REGION Network 25: Level Conveyors Tower 1 - SYSTEM 2
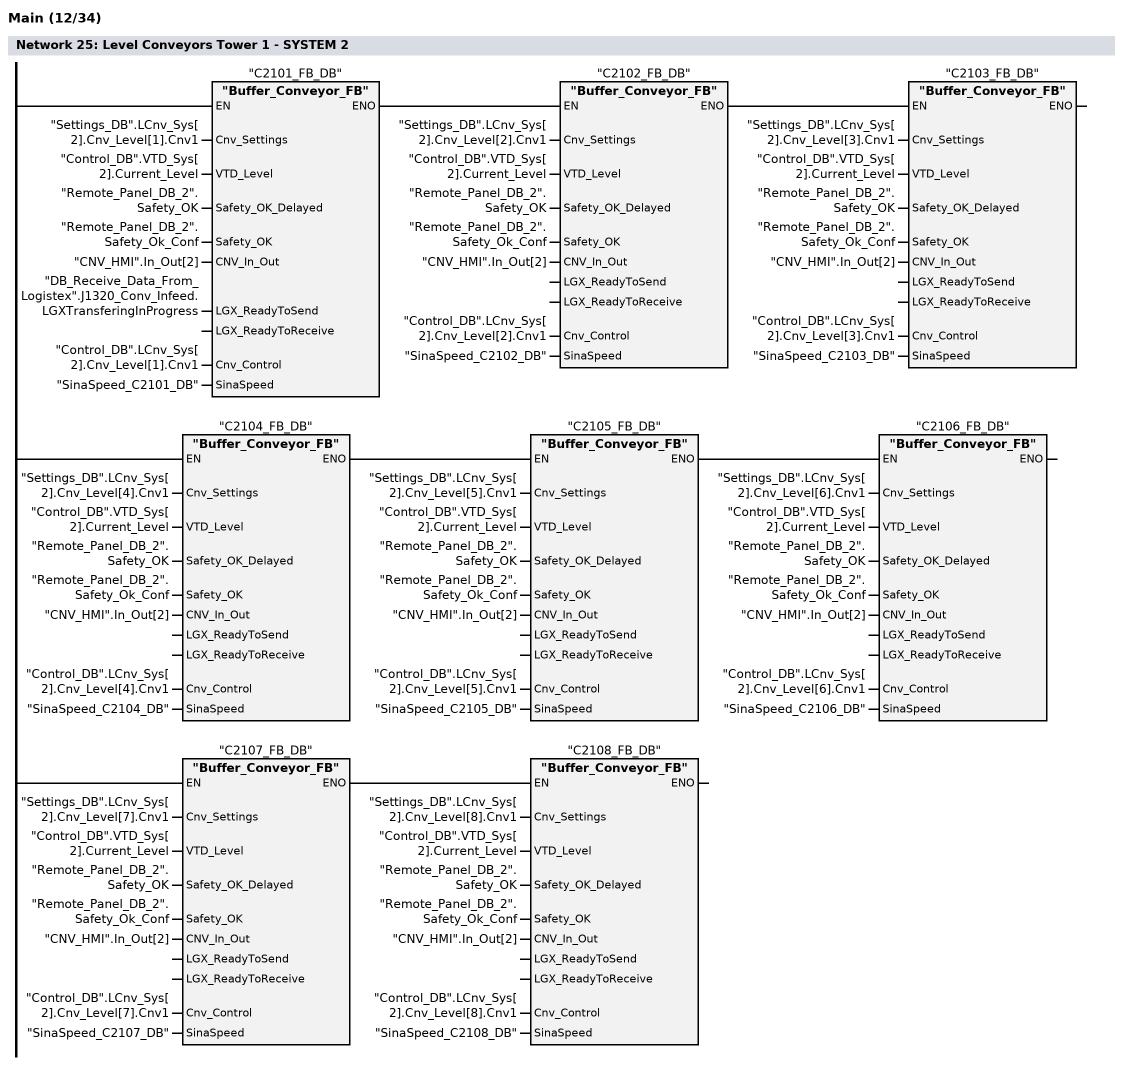
   RUNG wire#powerrail
      "C2101_FB_DB"(Cnv_Settings := "Settings_DB".LCnv_Sys[2].Cnv_Level[1].Cnv1, VTD_Level := "Control_DB".VTD_Sys[2].Current_Level, Safety_OK_Delayed := "Remote_Panel_DB_2".Safety_OK, Safety_OK := "Remote_Panel_DB_2".Safety_Ok_Conf, CNV_In_Out := "CNV_HMI".In_Out[2], LGX_ReadyToSend := "DB_Receive_Data_From_Logistex".J1320_Conv_Infeed.LGXTransferingInProgress, LGX_ReadyToReceive :=, Cnv_Control := "Control_DB".LCnv_Sys[2].Cnv_Level[1].Cnv1, SinaSpeed := "SinaSpeed_C2101_DB")
      "C2102_FB_DB"(Cnv_Settings := "Settings_DB".LCnv_Sys[2].Cnv_Level[2].Cnv1, VTD_Level := "Control_DB".VTD_Sys[2].Current_Level, Safety_OK_Delayed := "Remote_Panel_DB_2".Safety_OK, Safety_OK := "Remote_Panel_DB_2".Safety_Ok_Conf, CNV_In_Out := "CNV_HMI".In_Out[2], LGX_ReadyToSend :=, LGX_ReadyToReceive :=, Cnv_Control := "Control_DB".LCnv_Sys[2].Cnv_Level[2].Cnv1, SinaSpeed := "SinaSpeed_C2102_DB")
      "C2103_FB_DB"(Cnv_Settings := "Settings_DB".LCnv_Sys[2].Cnv_Level[3].Cnv1, VTD_Level := "Control_DB".VTD_Sys[2].Current_Level, Safety_OK_Delayed := "Remote_Panel_DB_2".Safety_OK, Safety_OK := "Remote_Panel_DB_2".Safety_Ok_Conf, CNV_In_Out := "CNV_HMI".In_Out[2], LGX_ReadyToSend :=, LGX_ReadyToReceive :=, Cnv_Control := "Control_DB".LCnv_Sys[2].Cnv_Level[3].Cnv1, SinaSpeed := "SinaSpeed_C2103_DB")
   END_RUNG
   RUNG wire#powerrail
      "C2104_FB_DB"(Cnv_Settings := "Settings_DB".LCnv_Sys[2].Cnv_Level[4].Cnv1, VTD_Level := "Control_DB".VTD_Sys[2].Current_Level, Safety_OK_Delayed := "Remote_Panel_DB_2".Safety_OK, Safety_OK := "Remote_Panel_DB_2".Safety_Ok_Conf, CNV_In_Out := "CNV_HMI".In_Out[2], LGX_ReadyToSend :=, LGX_ReadyToReceive :=, Cnv_Control := "Control_DB".LCnv_Sys[2].Cnv_Level[4].Cnv1, SinaSpeed := "SinaSpeed_C2104_DB")
      "C2105_FB_DB"(Cnv_Settings := "Settings_DB".LCnv_Sys[2].Cnv_Level[5].Cnv1, VTD_Level := "Control_DB".VTD_Sys[2].Current_Level, Safety_OK_Delayed := "Remote_Panel_DB_2".Safety_OK, Safety_OK := "Remote_Panel_DB_2".Safety_Ok_Conf, CNV_In_Out := "CNV_HMI".In_Out[2], LGX_ReadyToSend :=, LGX_ReadyToReceive :=, Cnv_Control := "Control_DB".LCnv_Sys[2].Cnv_Level[5].Cnv1, SinaSpeed := "SinaSpeed_C2105_DB")
      "C2106_FB_DB"(Cnv_Settings := "Settings_DB".LCnv_Sys[2].Cnv_Level[6].Cnv1, VTD_Level := "Control_DB".VTD_Sys[2].Current_Level, Safety_OK_Delayed := "Remote_Panel_DB_2".Safety_OK, Safety_OK := "Remote_Panel_DB_2".Safety_Ok_Conf, CNV_In_Out := "CNV_HMI".In_Out[2], LGX_ReadyToSend :=, LGX_ReadyToReceive :=, Cnv_Control := "Control_DB".LCnv_Sys[2].Cnv_Level[6].Cnv1, SinaSpeed := "SinaSpeed_C2106_DB")
   END_RUNG
   RUNG wire#powerrail
      "C2107_FB_DB"(Cnv_Settings := "Settings_DB".LCnv_Sys[2].Cnv_Level[7].Cnv1, VTD_Level := "Control_DB".VTD_Sys[2].Current_Level, Safety_OK_Delayed := "Remote_Panel_DB_2".Safety_OK, Safety_OK := "Remote_Panel_DB_2".Safety_Ok_Conf, CNV_In_Out := "CNV_HMI".In_Out[2], LGX_ReadyToSend :=, LGX_ReadyToReceive :=, Cnv_Control := "Control_DB".LCnv_Sys[2].Cnv_Level[7].Cnv1, SinaSpeed := "SinaSpeed_C2107_DB")
      "C2108_FB_DB"(Cnv_Settings := "Settings_DB".LCnv_Sys[2].Cnv_Level[8].Cnv1, VTD_Level := "Control_DB".VTD_Sys[2].Current_Level, Safety_OK_Delayed := "Remote_Panel_DB_2".Safety_OK, Safety_OK := "Remote_Panel_DB_2".Safety_Ok_Conf, CNV_In_Out := "CNV_HMI".In_Out[2], LGX_ReadyToSend :=, LGX_ReadyToReceive :=, Cnv_Control := "Control_DB".LCnv_Sys[2].Cnv_Level[8].Cnv1, SinaSpeed := "SinaSpeed_C2108_DB")
   END_RUNG
   // the same network as SCL:
   "C2101_FB_DB"(Cnv_Settings := "Settings_DB".LCnv_Sys[2].Cnv_Level[1].Cnv1,   // "Buffer_Conveyor_FB"
                 VTD_Level := "Control_DB".VTD_Sys[2].Current_Level,
                 Safety_OK_Delayed := "Remote_Panel_DB_2".Safety_OK,
                 Safety_OK := "Remote_Panel_DB_2".Safety_Ok_Conf,
                 CNV_In_Out := "CNV_HMI".In_Out[2],
                 LGX_ReadyToSend := "DB_Receive_Data_From_Logistex".J1320_Conv_Infeed.LGXTransferingInProgress,
                 Cnv_Control := "Control_DB".LCnv_Sys[2].Cnv_Level[1].Cnv1,
                 SinaSpeed := "SinaSpeed_C2101_DB",
                 ENO => #_w1);
   "C2102_FB_DB"(EN := #_w1,   // "Buffer_Conveyor_FB"
                 Cnv_Settings := "Settings_DB".LCnv_Sys[2].Cnv_Level[2].Cnv1,
                 VTD_Level := "Control_DB".VTD_Sys[2].Current_Level,
                 Safety_OK_Delayed := "Remote_Panel_DB_2".Safety_OK,
                 Safety_OK := "Remote_Panel_DB_2".Safety_Ok_Conf,
                 CNV_In_Out := "CNV_HMI".In_Out[2],
                 Cnv_Control := "Control_DB".LCnv_Sys[2].Cnv_Level[2].Cnv1,
                 SinaSpeed := "SinaSpeed_C2102_DB",
                 ENO => #_w2);
   IF #_w2 THEN
       "C2103_FB_DB"(Cnv_Settings := "Settings_DB".LCnv_Sys[2].Cnv_Level[3].Cnv1,   // "Buffer_Conveyor_FB"
                     VTD_Level := "Control_DB".VTD_Sys[2].Current_Level,
                     Safety_OK_Delayed := "Remote_Panel_DB_2".Safety_OK,
                     Safety_OK := "Remote_Panel_DB_2".Safety_Ok_Conf,
                     CNV_In_Out := "CNV_HMI".In_Out[2],
                     Cnv_Control := "Control_DB".LCnv_Sys[2].Cnv_Level[3].Cnv1,
                     SinaSpeed := "SinaSpeed_C2103_DB");
   END_IF;
   "C2104_FB_DB"(Cnv_Settings := "Settings_DB".LCnv_Sys[2].Cnv_Level[4].Cnv1,   // "Buffer_Conveyor_FB"
                 VTD_Level := "Control_DB".VTD_Sys[2].Current_Level,
                 Safety_OK_Delayed := "Remote_Panel_DB_2".Safety_OK,
                 Safety_OK := "Remote_Panel_DB_2".Safety_Ok_Conf,
                 CNV_In_Out := "CNV_HMI".In_Out[2],
                 Cnv_Control := "Control_DB".LCnv_Sys[2].Cnv_Level[4].Cnv1,
                 SinaSpeed := "SinaSpeed_C2104_DB",
                 ENO => #_w3);
   "C2105_FB_DB"(EN := #_w3,   // "Buffer_Conveyor_FB"
                 Cnv_Settings := "Settings_DB".LCnv_Sys[2].Cnv_Level[5].Cnv1,
                 VTD_Level := "Control_DB".VTD_Sys[2].Current_Level,
                 Safety_OK_Delayed := "Remote_Panel_DB_2".Safety_OK,
                 Safety_OK := "Remote_Panel_DB_2".Safety_Ok_Conf,
                 CNV_In_Out := "CNV_HMI".In_Out[2],
                 Cnv_Control := "Control_DB".LCnv_Sys[2].Cnv_Level[5].Cnv1,
                 SinaSpeed := "SinaSpeed_C2105_DB",
                 ENO => #_w4);
   IF #_w4 THEN
       "C2106_FB_DB"(Cnv_Settings := "Settings_DB".LCnv_Sys[2].Cnv_Level[6].Cnv1,   // "Buffer_Conveyor_FB"
                     VTD_Level := "Control_DB".VTD_Sys[2].Current_Level,
                     Safety_OK_Delayed := "Remote_Panel_DB_2".Safety_OK,
                     Safety_OK := "Remote_Panel_DB_2".Safety_Ok_Conf,
                     CNV_In_Out := "CNV_HMI".In_Out[2],
                     Cnv_Control := "Control_DB".LCnv_Sys[2].Cnv_Level[6].Cnv1,
                     SinaSpeed := "SinaSpeed_C2106_DB");
   END_IF;
   "C2107_FB_DB"(Cnv_Settings := "Settings_DB".LCnv_Sys[2].Cnv_Level[7].Cnv1,   // "Buffer_Conveyor_FB"
                 VTD_Level := "Control_DB".VTD_Sys[2].Current_Level,
                 Safety_OK_Delayed := "Remote_Panel_DB_2".Safety_OK,
                 Safety_OK := "Remote_Panel_DB_2".Safety_Ok_Conf,
                 CNV_In_Out := "CNV_HMI".In_Out[2],
                 Cnv_Control := "Control_DB".LCnv_Sys[2].Cnv_Level[7].Cnv1,
                 SinaSpeed := "SinaSpeed_C2107_DB",
                 ENO => #_w5);
   IF #_w5 THEN
       "C2108_FB_DB"(Cnv_Settings := "Settings_DB".LCnv_Sys[2].Cnv_Level[8].Cnv1,   // "Buffer_Conveyor_FB"
                     VTD_Level := "Control_DB".VTD_Sys[2].Current_Level,
                     Safety_OK_Delayed := "Remote_Panel_DB_2".Safety_OK,
                     Safety_OK := "Remote_Panel_DB_2".Safety_Ok_Conf,
                     CNV_In_Out := "CNV_HMI".In_Out[2],
                     Cnv_Control := "Control_DB".LCnv_Sys[2].Cnv_Level[8].Cnv1,
                     SinaSpeed := "SinaSpeed_C2108_DB");
   END_IF;
END_REGION

REGION Network 26: Level Conveyors Tower 2 - SYSTEM 2
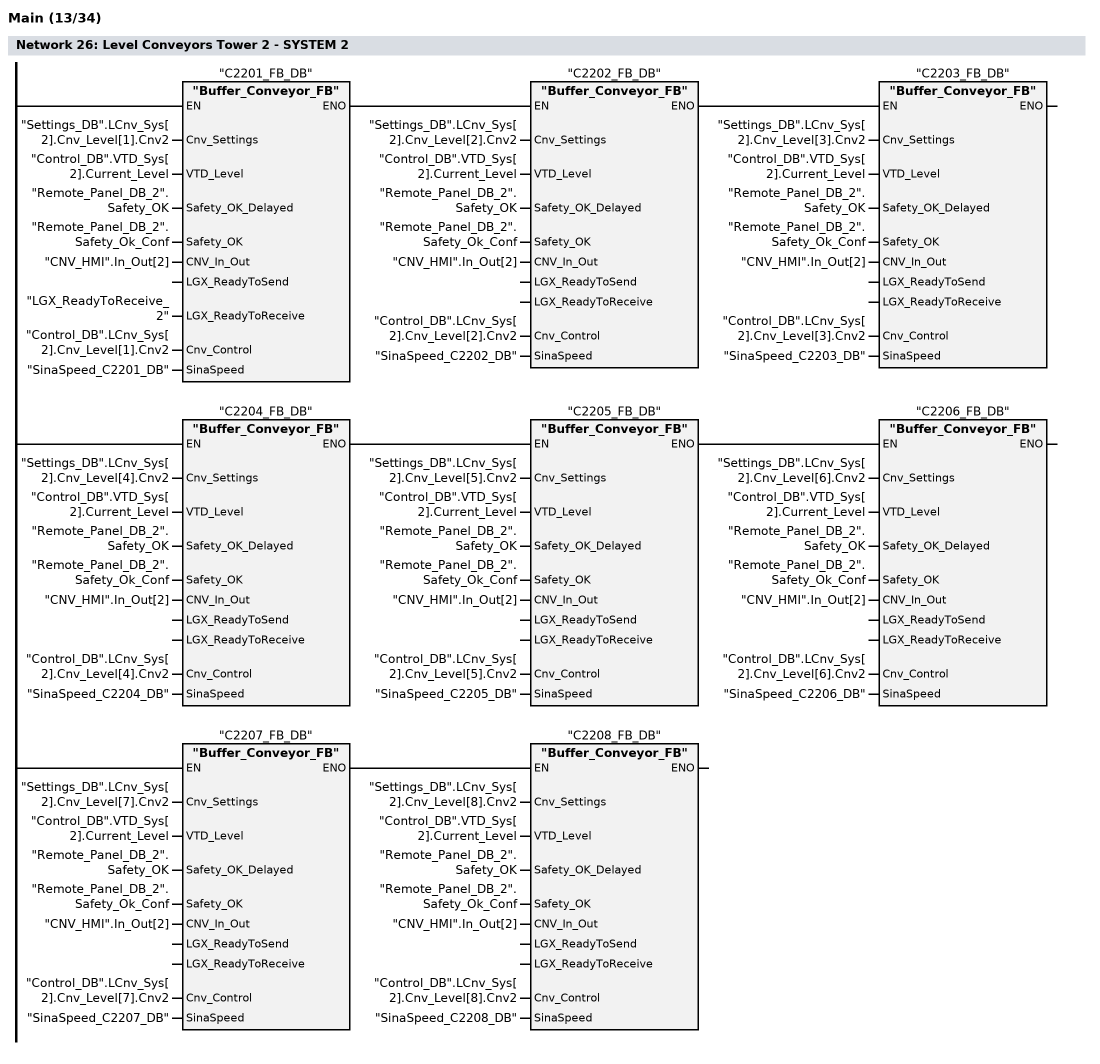
   RUNG wire#powerrail
      "C2201_FB_DB"(Cnv_Settings := "Settings_DB".LCnv_Sys[2].Cnv_Level[1].Cnv2, VTD_Level := "Control_DB".VTD_Sys[2].Current_Level, Safety_OK_Delayed := "Remote_Panel_DB_2".Safety_OK, Safety_OK := "Remote_Panel_DB_2".Safety_Ok_Conf, CNV_In_Out := "CNV_HMI".In_Out[2], LGX_ReadyToSend :=, LGX_ReadyToReceive := "LGX_ReadyToReceive_2", Cnv_Control := "Control_DB".LCnv_Sys[2].Cnv_Level[1].Cnv2, SinaSpeed := "SinaSpeed_C2201_DB")
      "C2202_FB_DB"(Cnv_Settings := "Settings_DB".LCnv_Sys[2].Cnv_Level[2].Cnv2, VTD_Level := "Control_DB".VTD_Sys[2].Current_Level, Safety_OK_Delayed := "Remote_Panel_DB_2".Safety_OK, Safety_OK := "Remote_Panel_DB_2".Safety_Ok_Conf, CNV_In_Out := "CNV_HMI".In_Out[2], LGX_ReadyToSend :=, LGX_ReadyToReceive :=, Cnv_Control := "Control_DB".LCnv_Sys[2].Cnv_Level[2].Cnv2, SinaSpeed := "SinaSpeed_C2202_DB")
      "C2203_FB_DB"(Cnv_Settings := "Settings_DB".LCnv_Sys[2].Cnv_Level[3].Cnv2, VTD_Level := "Control_DB".VTD_Sys[2].Current_Level, Safety_OK_Delayed := "Remote_Panel_DB_2".Safety_OK, Safety_OK := "Remote_Panel_DB_2".Safety_Ok_Conf, CNV_In_Out := "CNV_HMI".In_Out[2], LGX_ReadyToSend :=, LGX_ReadyToReceive :=, Cnv_Control := "Control_DB".LCnv_Sys[2].Cnv_Level[3].Cnv2, SinaSpeed := "SinaSpeed_C2203_DB")
   END_RUNG
   RUNG wire#powerrail
      "C2204_FB_DB"(Cnv_Settings := "Settings_DB".LCnv_Sys[2].Cnv_Level[4].Cnv2, VTD_Level := "Control_DB".VTD_Sys[2].Current_Level, Safety_OK_Delayed := "Remote_Panel_DB_2".Safety_OK, Safety_OK := "Remote_Panel_DB_2".Safety_Ok_Conf, CNV_In_Out := "CNV_HMI".In_Out[2], LGX_ReadyToSend :=, LGX_ReadyToReceive :=, Cnv_Control := "Control_DB".LCnv_Sys[2].Cnv_Level[4].Cnv2, SinaSpeed := "SinaSpeed_C2204_DB")
      "C2205_FB_DB"(Cnv_Settings := "Settings_DB".LCnv_Sys[2].Cnv_Level[5].Cnv2, VTD_Level := "Control_DB".VTD_Sys[2].Current_Level, Safety_OK_Delayed := "Remote_Panel_DB_2".Safety_OK, Safety_OK := "Remote_Panel_DB_2".Safety_Ok_Conf, CNV_In_Out := "CNV_HMI".In_Out[2], LGX_ReadyToSend :=, LGX_ReadyToReceive :=, Cnv_Control := "Control_DB".LCnv_Sys[2].Cnv_Level[5].Cnv2, SinaSpeed := "SinaSpeed_C2205_DB")
      "C2206_FB_DB"(Cnv_Settings := "Settings_DB".LCnv_Sys[2].Cnv_Level[6].Cnv2, VTD_Level := "Control_DB".VTD_Sys[2].Current_Level, Safety_OK_Delayed := "Remote_Panel_DB_2".Safety_OK, Safety_OK := "Remote_Panel_DB_2".Safety_Ok_Conf, CNV_In_Out := "CNV_HMI".In_Out[2], LGX_ReadyToSend :=, LGX_ReadyToReceive :=, Cnv_Control := "Control_DB".LCnv_Sys[2].Cnv_Level[6].Cnv2, SinaSpeed := "SinaSpeed_C2206_DB")
   END_RUNG
   RUNG wire#powerrail
      "C2207_FB_DB"(Cnv_Settings := "Settings_DB".LCnv_Sys[2].Cnv_Level[7].Cnv2, VTD_Level := "Control_DB".VTD_Sys[2].Current_Level, Safety_OK_Delayed := "Remote_Panel_DB_2".Safety_OK, Safety_OK := "Remote_Panel_DB_2".Safety_Ok_Conf, CNV_In_Out := "CNV_HMI".In_Out[2], LGX_ReadyToSend :=, LGX_ReadyToReceive :=, Cnv_Control := "Control_DB".LCnv_Sys[2].Cnv_Level[7].Cnv2, SinaSpeed := "SinaSpeed_C2207_DB")
      "C2208_FB_DB"(Cnv_Settings := "Settings_DB".LCnv_Sys[2].Cnv_Level[8].Cnv2, VTD_Level := "Control_DB".VTD_Sys[2].Current_Level, Safety_OK_Delayed := "Remote_Panel_DB_2".Safety_OK, Safety_OK := "Remote_Panel_DB_2".Safety_Ok_Conf, CNV_In_Out := "CNV_HMI".In_Out[2], LGX_ReadyToSend :=, LGX_ReadyToReceive :=, Cnv_Control := "Control_DB".LCnv_Sys[2].Cnv_Level[8].Cnv2, SinaSpeed := "SinaSpeed_C2208_DB")
   END_RUNG
   // the same network as SCL:
   "C2201_FB_DB"(Cnv_Settings := "Settings_DB".LCnv_Sys[2].Cnv_Level[1].Cnv2,   // "Buffer_Conveyor_FB"
                 VTD_Level := "Control_DB".VTD_Sys[2].Current_Level,
                 Safety_OK_Delayed := "Remote_Panel_DB_2".Safety_OK,
                 Safety_OK := "Remote_Panel_DB_2".Safety_Ok_Conf,
                 CNV_In_Out := "CNV_HMI".In_Out[2],
                 LGX_ReadyToReceive := "LGX_ReadyToReceive_2",
                 Cnv_Control := "Control_DB".LCnv_Sys[2].Cnv_Level[1].Cnv2,
                 SinaSpeed := "SinaSpeed_C2201_DB",
                 ENO => #_w1);
   "C2202_FB_DB"(EN := #_w1,   // "Buffer_Conveyor_FB"
                 Cnv_Settings := "Settings_DB".LCnv_Sys[2].Cnv_Level[2].Cnv2,
                 VTD_Level := "Control_DB".VTD_Sys[2].Current_Level,
                 Safety_OK_Delayed := "Remote_Panel_DB_2".Safety_OK,
                 Safety_OK := "Remote_Panel_DB_2".Safety_Ok_Conf,
                 CNV_In_Out := "CNV_HMI".In_Out[2],
                 Cnv_Control := "Control_DB".LCnv_Sys[2].Cnv_Level[2].Cnv2,
                 SinaSpeed := "SinaSpeed_C2202_DB",
                 ENO => #_w2);
   IF #_w2 THEN
       "C2203_FB_DB"(Cnv_Settings := "Settings_DB".LCnv_Sys[2].Cnv_Level[3].Cnv2,   // "Buffer_Conveyor_FB"
                     VTD_Level := "Control_DB".VTD_Sys[2].Current_Level,
                     Safety_OK_Delayed := "Remote_Panel_DB_2".Safety_OK,
                     Safety_OK := "Remote_Panel_DB_2".Safety_Ok_Conf,
                     CNV_In_Out := "CNV_HMI".In_Out[2],
                     Cnv_Control := "Control_DB".LCnv_Sys[2].Cnv_Level[3].Cnv2,
                     SinaSpeed := "SinaSpeed_C2203_DB");
   END_IF;
   "C2204_FB_DB"(Cnv_Settings := "Settings_DB".LCnv_Sys[2].Cnv_Level[4].Cnv2,   // "Buffer_Conveyor_FB"
                 VTD_Level := "Control_DB".VTD_Sys[2].Current_Level,
                 Safety_OK_Delayed := "Remote_Panel_DB_2".Safety_OK,
                 Safety_OK := "Remote_Panel_DB_2".Safety_Ok_Conf,
                 CNV_In_Out := "CNV_HMI".In_Out[2],
                 Cnv_Control := "Control_DB".LCnv_Sys[2].Cnv_Level[4].Cnv2,
                 SinaSpeed := "SinaSpeed_C2204_DB",
                 ENO => #_w3);
   "C2205_FB_DB"(EN := #_w3,   // "Buffer_Conveyor_FB"
                 Cnv_Settings := "Settings_DB".LCnv_Sys[2].Cnv_Level[5].Cnv2,
                 VTD_Level := "Control_DB".VTD_Sys[2].Current_Level,
                 Safety_OK_Delayed := "Remote_Panel_DB_2".Safety_OK,
                 Safety_OK := "Remote_Panel_DB_2".Safety_Ok_Conf,
                 CNV_In_Out := "CNV_HMI".In_Out[2],
                 Cnv_Control := "Control_DB".LCnv_Sys[2].Cnv_Level[5].Cnv2,
                 SinaSpeed := "SinaSpeed_C2205_DB",
                 ENO => #_w4);
   IF #_w4 THEN
       "C2206_FB_DB"(Cnv_Settings := "Settings_DB".LCnv_Sys[2].Cnv_Level[6].Cnv2,   // "Buffer_Conveyor_FB"
                     VTD_Level := "Control_DB".VTD_Sys[2].Current_Level,
                     Safety_OK_Delayed := "Remote_Panel_DB_2".Safety_OK,
                     Safety_OK := "Remote_Panel_DB_2".Safety_Ok_Conf,
                     CNV_In_Out := "CNV_HMI".In_Out[2],
                     Cnv_Control := "Control_DB".LCnv_Sys[2].Cnv_Level[6].Cnv2,
                     SinaSpeed := "SinaSpeed_C2206_DB");
   END_IF;
   "C2207_FB_DB"(Cnv_Settings := "Settings_DB".LCnv_Sys[2].Cnv_Level[7].Cnv2,   // "Buffer_Conveyor_FB"
                 VTD_Level := "Control_DB".VTD_Sys[2].Current_Level,
                 Safety_OK_Delayed := "Remote_Panel_DB_2".Safety_OK,
                 Safety_OK := "Remote_Panel_DB_2".Safety_Ok_Conf,
                 CNV_In_Out := "CNV_HMI".In_Out[2],
                 Cnv_Control := "Control_DB".LCnv_Sys[2].Cnv_Level[7].Cnv2,
                 SinaSpeed := "SinaSpeed_C2207_DB",
                 ENO => #_w5);
   IF #_w5 THEN
       "C2208_FB_DB"(Cnv_Settings := "Settings_DB".LCnv_Sys[2].Cnv_Level[8].Cnv2,   // "Buffer_Conveyor_FB"
                     VTD_Level := "Control_DB".VTD_Sys[2].Current_Level,
                     Safety_OK_Delayed := "Remote_Panel_DB_2".Safety_OK,
                     Safety_OK := "Remote_Panel_DB_2".Safety_Ok_Conf,
                     CNV_In_Out := "CNV_HMI".In_Out[2],
                     Cnv_Control := "Control_DB".LCnv_Sys[2].Cnv_Level[8].Cnv2,
                     SinaSpeed := "SinaSpeed_C2208_DB");
   END_IF;
END_REGION

REGION Network 27: SAFETY STOPPERS Tower 1 - SYSTEM 2
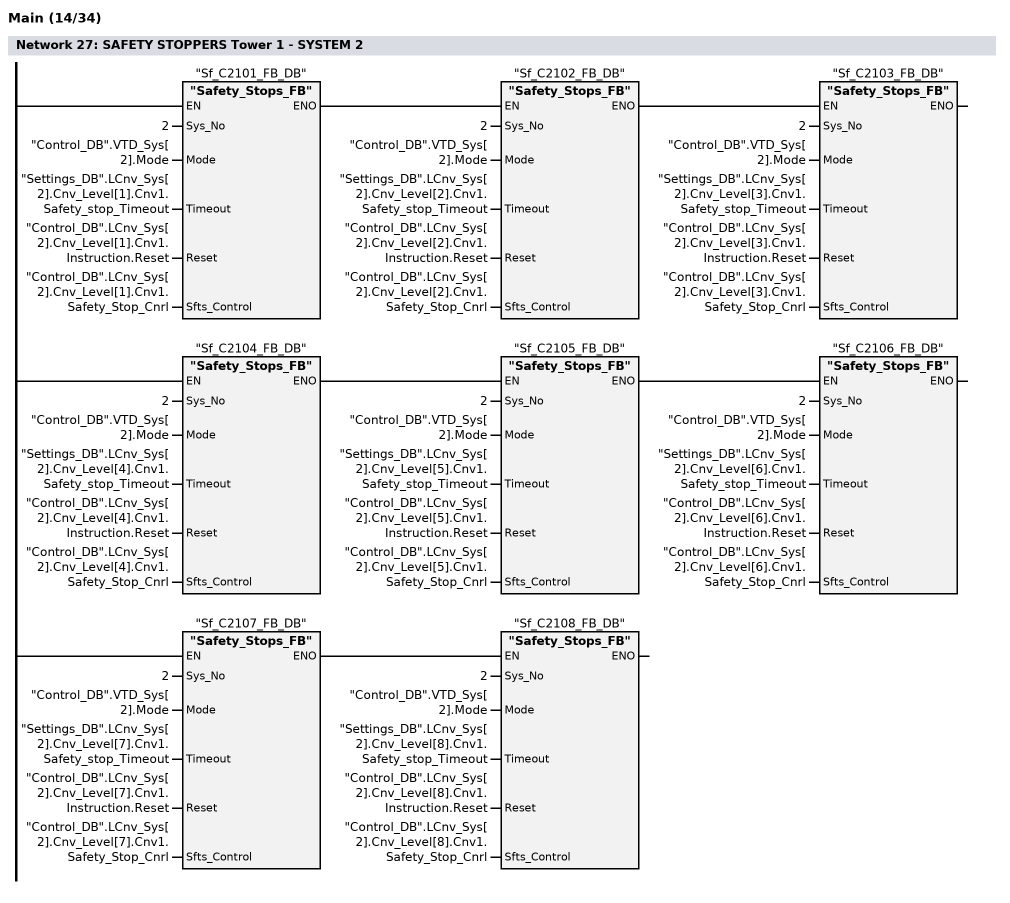
   RUNG wire#powerrail
      "Sf_C2101_FB_DB"(Sys_No := 2, Mode := "Control_DB".VTD_Sys[2].Mode, Timeout := "Settings_DB".LCnv_Sys[2].Cnv_Level[1].Cnv1.Safety_stop_Timeout, Reset := "Control_DB".LCnv_Sys[2].Cnv_Level[1].Cnv1.Instruction.Reset, Sfts_Control := "Control_DB".LCnv_Sys[2].Cnv_Level[1].Cnv1.Safety_Stop_Cnrl)
      "Sf_C2102_FB_DB"(Sys_No := 2, Mode := "Control_DB".VTD_Sys[2].Mode, Timeout := "Settings_DB".LCnv_Sys[2].Cnv_Level[2].Cnv1.Safety_stop_Timeout, Reset := "Control_DB".LCnv_Sys[2].Cnv_Level[2].Cnv1.Instruction.Reset, Sfts_Control := "Control_DB".LCnv_Sys[2].Cnv_Level[2].Cnv1.Safety_Stop_Cnrl)
      "Sf_C2103_FB_DB"(Sys_No := 2, Mode := "Control_DB".VTD_Sys[2].Mode, Timeout := "Settings_DB".LCnv_Sys[2].Cnv_Level[3].Cnv1.Safety_stop_Timeout, Reset := "Control_DB".LCnv_Sys[2].Cnv_Level[3].Cnv1.Instruction.Reset, Sfts_Control := "Control_DB".LCnv_Sys[2].Cnv_Level[3].Cnv1.Safety_Stop_Cnrl)
   END_RUNG
   RUNG wire#powerrail
      "Sf_C2104_FB_DB"(Sys_No := 2, Mode := "Control_DB".VTD_Sys[2].Mode, Timeout := "Settings_DB".LCnv_Sys[2].Cnv_Level[4].Cnv1.Safety_stop_Timeout, Reset := "Control_DB".LCnv_Sys[2].Cnv_Level[4].Cnv1.Instruction.Reset, Sfts_Control := "Control_DB".LCnv_Sys[2].Cnv_Level[4].Cnv1.Safety_Stop_Cnrl)
      "Sf_C2105_FB_DB"(Sys_No := 2, Mode := "Control_DB".VTD_Sys[2].Mode, Timeout := "Settings_DB".LCnv_Sys[2].Cnv_Level[5].Cnv1.Safety_stop_Timeout, Reset := "Control_DB".LCnv_Sys[2].Cnv_Level[5].Cnv1.Instruction.Reset, Sfts_Control := "Control_DB".LCnv_Sys[2].Cnv_Level[5].Cnv1.Safety_Stop_Cnrl)
      "Sf_C2106_FB_DB"(Sys_No := 2, Mode := "Control_DB".VTD_Sys[2].Mode, Timeout := "Settings_DB".LCnv_Sys[2].Cnv_Level[6].Cnv1.Safety_stop_Timeout, Reset := "Control_DB".LCnv_Sys[2].Cnv_Level[6].Cnv1.Instruction.Reset, Sfts_Control := "Control_DB".LCnv_Sys[2].Cnv_Level[6].Cnv1.Safety_Stop_Cnrl)
   END_RUNG
   RUNG wire#powerrail
      "Sf_C2107_FB_DB"(Sys_No := 2, Mode := "Control_DB".VTD_Sys[2].Mode, Timeout := "Settings_DB".LCnv_Sys[2].Cnv_Level[7].Cnv1.Safety_stop_Timeout, Reset := "Control_DB".LCnv_Sys[2].Cnv_Level[7].Cnv1.Instruction.Reset, Sfts_Control := "Control_DB".LCnv_Sys[2].Cnv_Level[7].Cnv1.Safety_Stop_Cnrl)
      "Sf_C2108_FB_DB"(Sys_No := 2, Mode := "Control_DB".VTD_Sys[2].Mode, Timeout := "Settings_DB".LCnv_Sys[2].Cnv_Level[8].Cnv1.Safety_stop_Timeout, Reset := "Control_DB".LCnv_Sys[2].Cnv_Level[8].Cnv1.Instruction.Reset, Sfts_Control := "Control_DB".LCnv_Sys[2].Cnv_Level[8].Cnv1.Safety_Stop_Cnrl)
   END_RUNG
   // the same network as SCL:
   "Sf_C2101_FB_DB"(Sys_No := 2,   // "Safety_Stops_FB"
                    Mode := "Control_DB".VTD_Sys[2].Mode,
                    Timeout := "Settings_DB".LCnv_Sys[2].Cnv_Level[1].Cnv1.Safety_stop_Timeout,
                    Reset := "Control_DB".LCnv_Sys[2].Cnv_Level[1].Cnv1.Instruction.Reset,
                    Sfts_Control := "Control_DB".LCnv_Sys[2].Cnv_Level[1].Cnv1.Safety_Stop_Cnrl,
                    ENO => #_w1);
   "Sf_C2102_FB_DB"(EN := #_w1,   // "Safety_Stops_FB"
                    Sys_No := 2,
                    Mode := "Control_DB".VTD_Sys[2].Mode,
                    Timeout := "Settings_DB".LCnv_Sys[2].Cnv_Level[2].Cnv1.Safety_stop_Timeout,
                    Reset := "Control_DB".LCnv_Sys[2].Cnv_Level[2].Cnv1.Instruction.Reset,
                    Sfts_Control := "Control_DB".LCnv_Sys[2].Cnv_Level[2].Cnv1.Safety_Stop_Cnrl,
                    ENO => #_w2);
   IF #_w2 THEN
       "Sf_C2103_FB_DB"(Sys_No := 2,   // "Safety_Stops_FB"
                        Mode := "Control_DB".VTD_Sys[2].Mode,
                        Timeout := "Settings_DB".LCnv_Sys[2].Cnv_Level[3].Cnv1.Safety_stop_Timeout,
                        Reset := "Control_DB".LCnv_Sys[2].Cnv_Level[3].Cnv1.Instruction.Reset,
                        Sfts_Control := "Control_DB".LCnv_Sys[2].Cnv_Level[3].Cnv1.Safety_Stop_Cnrl);
   END_IF;
   "Sf_C2104_FB_DB"(Sys_No := 2,   // "Safety_Stops_FB"
                    Mode := "Control_DB".VTD_Sys[2].Mode,
                    Timeout := "Settings_DB".LCnv_Sys[2].Cnv_Level[4].Cnv1.Safety_stop_Timeout,
                    Reset := "Control_DB".LCnv_Sys[2].Cnv_Level[4].Cnv1.Instruction.Reset,
                    Sfts_Control := "Control_DB".LCnv_Sys[2].Cnv_Level[4].Cnv1.Safety_Stop_Cnrl,
                    ENO => #_w3);
   "Sf_C2105_FB_DB"(EN := #_w3,   // "Safety_Stops_FB"
                    Sys_No := 2,
                    Mode := "Control_DB".VTD_Sys[2].Mode,
                    Timeout := "Settings_DB".LCnv_Sys[2].Cnv_Level[5].Cnv1.Safety_stop_Timeout,
                    Reset := "Control_DB".LCnv_Sys[2].Cnv_Level[5].Cnv1.Instruction.Reset,
                    Sfts_Control := "Control_DB".LCnv_Sys[2].Cnv_Level[5].Cnv1.Safety_Stop_Cnrl,
                    ENO => #_w4);
   IF #_w4 THEN
       "Sf_C2106_FB_DB"(Sys_No := 2,   // "Safety_Stops_FB"
                        Mode := "Control_DB".VTD_Sys[2].Mode,
                        Timeout := "Settings_DB".LCnv_Sys[2].Cnv_Level[6].Cnv1.Safety_stop_Timeout,
                        Reset := "Control_DB".LCnv_Sys[2].Cnv_Level[6].Cnv1.Instruction.Reset,
                        Sfts_Control := "Control_DB".LCnv_Sys[2].Cnv_Level[6].Cnv1.Safety_Stop_Cnrl);
   END_IF;
   "Sf_C2107_FB_DB"(Sys_No := 2,   // "Safety_Stops_FB"
                    Mode := "Control_DB".VTD_Sys[2].Mode,
                    Timeout := "Settings_DB".LCnv_Sys[2].Cnv_Level[7].Cnv1.Safety_stop_Timeout,
                    Reset := "Control_DB".LCnv_Sys[2].Cnv_Level[7].Cnv1.Instruction.Reset,
                    Sfts_Control := "Control_DB".LCnv_Sys[2].Cnv_Level[7].Cnv1.Safety_Stop_Cnrl,
                    ENO => #_w5);
   IF #_w5 THEN
       "Sf_C2108_FB_DB"(Sys_No := 2,   // "Safety_Stops_FB"
                        Mode := "Control_DB".VTD_Sys[2].Mode,
                        Timeout := "Settings_DB".LCnv_Sys[2].Cnv_Level[8].Cnv1.Safety_stop_Timeout,
                        Reset := "Control_DB".LCnv_Sys[2].Cnv_Level[8].Cnv1.Instruction.Reset,
                        Sfts_Control := "Control_DB".LCnv_Sys[2].Cnv_Level[8].Cnv1.Safety_Stop_Cnrl);
   END_IF;
END_REGION

REGION Network 28: SAFETY STOPPERS Tower 2 - SYSTEM 2
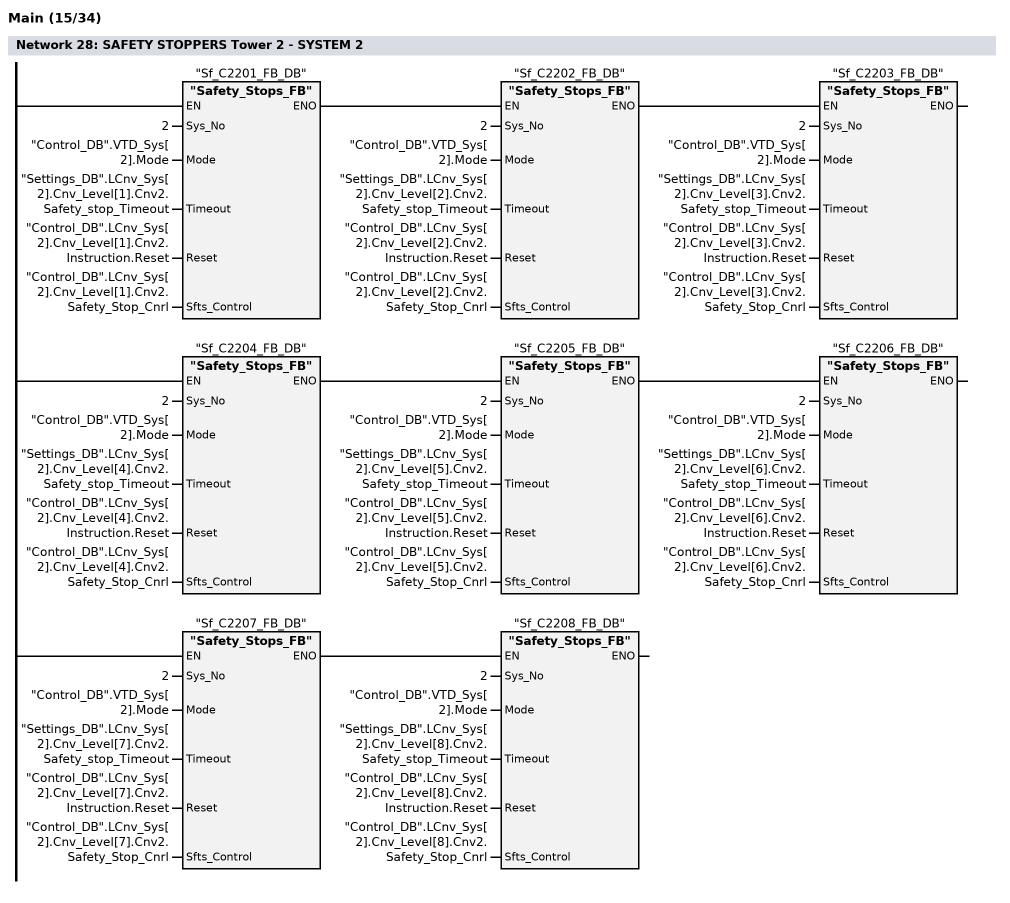
   RUNG wire#powerrail
      "Sf_C2201_FB_DB"(Sys_No := 2, Mode := "Control_DB".VTD_Sys[2].Mode, Timeout := "Settings_DB".LCnv_Sys[2].Cnv_Level[1].Cnv2.Safety_stop_Timeout, Reset := "Control_DB".LCnv_Sys[2].Cnv_Level[1].Cnv2.Instruction.Reset, Sfts_Control := "Control_DB".LCnv_Sys[2].Cnv_Level[1].Cnv2.Safety_Stop_Cnrl)
      "Sf_C2202_FB_DB"(Sys_No := 2, Mode := "Control_DB".VTD_Sys[2].Mode, Timeout := "Settings_DB".LCnv_Sys[2].Cnv_Level[2].Cnv2.Safety_stop_Timeout, Reset := "Control_DB".LCnv_Sys[2].Cnv_Level[2].Cnv2.Instruction.Reset, Sfts_Control := "Control_DB".LCnv_Sys[2].Cnv_Level[2].Cnv2.Safety_Stop_Cnrl)
      "Sf_C2203_FB_DB"(Sys_No := 2, Mode := "Control_DB".VTD_Sys[2].Mode, Timeout := "Settings_DB".LCnv_Sys[2].Cnv_Level[3].Cnv2.Safety_stop_Timeout, Reset := "Control_DB".LCnv_Sys[2].Cnv_Level[3].Cnv2.Instruction.Reset, Sfts_Control := "Control_DB".LCnv_Sys[2].Cnv_Level[3].Cnv2.Safety_Stop_Cnrl)
   END_RUNG
   RUNG wire#powerrail
      "Sf_C2204_FB_DB"(Sys_No := 2, Mode := "Control_DB".VTD_Sys[2].Mode, Timeout := "Settings_DB".LCnv_Sys[2].Cnv_Level[4].Cnv2.Safety_stop_Timeout, Reset := "Control_DB".LCnv_Sys[2].Cnv_Level[4].Cnv2.Instruction.Reset, Sfts_Control := "Control_DB".LCnv_Sys[2].Cnv_Level[4].Cnv2.Safety_Stop_Cnrl)
      "Sf_C2205_FB_DB"(Sys_No := 2, Mode := "Control_DB".VTD_Sys[2].Mode, Timeout := "Settings_DB".LCnv_Sys[2].Cnv_Level[5].Cnv2.Safety_stop_Timeout, Reset := "Control_DB".LCnv_Sys[2].Cnv_Level[5].Cnv2.Instruction.Reset, Sfts_Control := "Control_DB".LCnv_Sys[2].Cnv_Level[5].Cnv2.Safety_Stop_Cnrl)
      "Sf_C2206_FB_DB"(Sys_No := 2, Mode := "Control_DB".VTD_Sys[2].Mode, Timeout := "Settings_DB".LCnv_Sys[2].Cnv_Level[6].Cnv2.Safety_stop_Timeout, Reset := "Control_DB".LCnv_Sys[2].Cnv_Level[6].Cnv2.Instruction.Reset, Sfts_Control := "Control_DB".LCnv_Sys[2].Cnv_Level[6].Cnv2.Safety_Stop_Cnrl)
   END_RUNG
   RUNG wire#powerrail
      "Sf_C2207_FB_DB"(Sys_No := 2, Mode := "Control_DB".VTD_Sys[2].Mode, Timeout := "Settings_DB".LCnv_Sys[2].Cnv_Level[7].Cnv2.Safety_stop_Timeout, Reset := "Control_DB".LCnv_Sys[2].Cnv_Level[7].Cnv2.Instruction.Reset, Sfts_Control := "Control_DB".LCnv_Sys[2].Cnv_Level[7].Cnv2.Safety_Stop_Cnrl)
      "Sf_C2208_FB_DB"(Sys_No := 2, Mode := "Control_DB".VTD_Sys[2].Mode, Timeout := "Settings_DB".LCnv_Sys[2].Cnv_Level[8].Cnv2.Safety_stop_Timeout, Reset := "Control_DB".LCnv_Sys[2].Cnv_Level[8].Cnv2.Instruction.Reset, Sfts_Control := "Control_DB".LCnv_Sys[2].Cnv_Level[8].Cnv2.Safety_Stop_Cnrl)
   END_RUNG
   // the same network as SCL:
   "Sf_C2201_FB_DB"(Sys_No := 2,   // "Safety_Stops_FB"
                    Mode := "Control_DB".VTD_Sys[2].Mode,
                    Timeout := "Settings_DB".LCnv_Sys[2].Cnv_Level[1].Cnv2.Safety_stop_Timeout,
                    Reset := "Control_DB".LCnv_Sys[2].Cnv_Level[1].Cnv2.Instruction.Reset,
                    Sfts_Control := "Control_DB".LCnv_Sys[2].Cnv_Level[1].Cnv2.Safety_Stop_Cnrl,
                    ENO => #_w1);
   "Sf_C2202_FB_DB"(EN := #_w1,   // "Safety_Stops_FB"
                    Sys_No := 2,
                    Mode := "Control_DB".VTD_Sys[2].Mode,
                    Timeout := "Settings_DB".LCnv_Sys[2].Cnv_Level[2].Cnv2.Safety_stop_Timeout,
                    Reset := "Control_DB".LCnv_Sys[2].Cnv_Level[2].Cnv2.Instruction.Reset,
                    Sfts_Control := "Control_DB".LCnv_Sys[2].Cnv_Level[2].Cnv2.Safety_Stop_Cnrl,
                    ENO => #_w2);
   IF #_w2 THEN
       "Sf_C2203_FB_DB"(Sys_No := 2,   // "Safety_Stops_FB"
                        Mode := "Control_DB".VTD_Sys[2].Mode,
                        Timeout := "Settings_DB".LCnv_Sys[2].Cnv_Level[3].Cnv2.Safety_stop_Timeout,
                        Reset := "Control_DB".LCnv_Sys[2].Cnv_Level[3].Cnv2.Instruction.Reset,
                        Sfts_Control := "Control_DB".LCnv_Sys[2].Cnv_Level[3].Cnv2.Safety_Stop_Cnrl);
   END_IF;
   "Sf_C2204_FB_DB"(Sys_No := 2,   // "Safety_Stops_FB"
                    Mode := "Control_DB".VTD_Sys[2].Mode,
                    Timeout := "Settings_DB".LCnv_Sys[2].Cnv_Level[4].Cnv2.Safety_stop_Timeout,
                    Reset := "Control_DB".LCnv_Sys[2].Cnv_Level[4].Cnv2.Instruction.Reset,
                    Sfts_Control := "Control_DB".LCnv_Sys[2].Cnv_Level[4].Cnv2.Safety_Stop_Cnrl,
                    ENO => #_w3);
   "Sf_C2205_FB_DB"(EN := #_w3,   // "Safety_Stops_FB"
                    Sys_No := 2,
                    Mode := "Control_DB".VTD_Sys[2].Mode,
                    Timeout := "Settings_DB".LCnv_Sys[2].Cnv_Level[5].Cnv2.Safety_stop_Timeout,
                    Reset := "Control_DB".LCnv_Sys[2].Cnv_Level[5].Cnv2.Instruction.Reset,
                    Sfts_Control := "Control_DB".LCnv_Sys[2].Cnv_Level[5].Cnv2.Safety_Stop_Cnrl,
                    ENO => #_w4);
   IF #_w4 THEN
       "Sf_C2206_FB_DB"(Sys_No := 2,   // "Safety_Stops_FB"
                        Mode := "Control_DB".VTD_Sys[2].Mode,
                        Timeout := "Settings_DB".LCnv_Sys[2].Cnv_Level[6].Cnv2.Safety_stop_Timeout,
                        Reset := "Control_DB".LCnv_Sys[2].Cnv_Level[6].Cnv2.Instruction.Reset,
                        Sfts_Control := "Control_DB".LCnv_Sys[2].Cnv_Level[6].Cnv2.Safety_Stop_Cnrl);
   END_IF;
   "Sf_C2207_FB_DB"(Sys_No := 2,   // "Safety_Stops_FB"
                    Mode := "Control_DB".VTD_Sys[2].Mode,
                    Timeout := "Settings_DB".LCnv_Sys[2].Cnv_Level[7].Cnv2.Safety_stop_Timeout,
                    Reset := "Control_DB".LCnv_Sys[2].Cnv_Level[7].Cnv2.Instruction.Reset,
                    Sfts_Control := "Control_DB".LCnv_Sys[2].Cnv_Level[7].Cnv2.Safety_Stop_Cnrl,
                    ENO => #_w5);
   IF #_w5 THEN
       "Sf_C2208_FB_DB"(Sys_No := 2,   // "Safety_Stops_FB"
                        Mode := "Control_DB".VTD_Sys[2].Mode,
                        Timeout := "Settings_DB".LCnv_Sys[2].Cnv_Level[8].Cnv2.Safety_stop_Timeout,
                        Reset := "Control_DB".LCnv_Sys[2].Cnv_Level[8].Cnv2.Instruction.Reset,
                        Sfts_Control := "Control_DB".LCnv_Sys[2].Cnv_Level[8].Cnv2.Safety_Stop_Cnrl);
   END_IF;
END_REGION

REGION Network 29: SYSTEM 3
END_REGION

REGION Network 30: Level Conveyors Tower 1 - SYSTEM 3
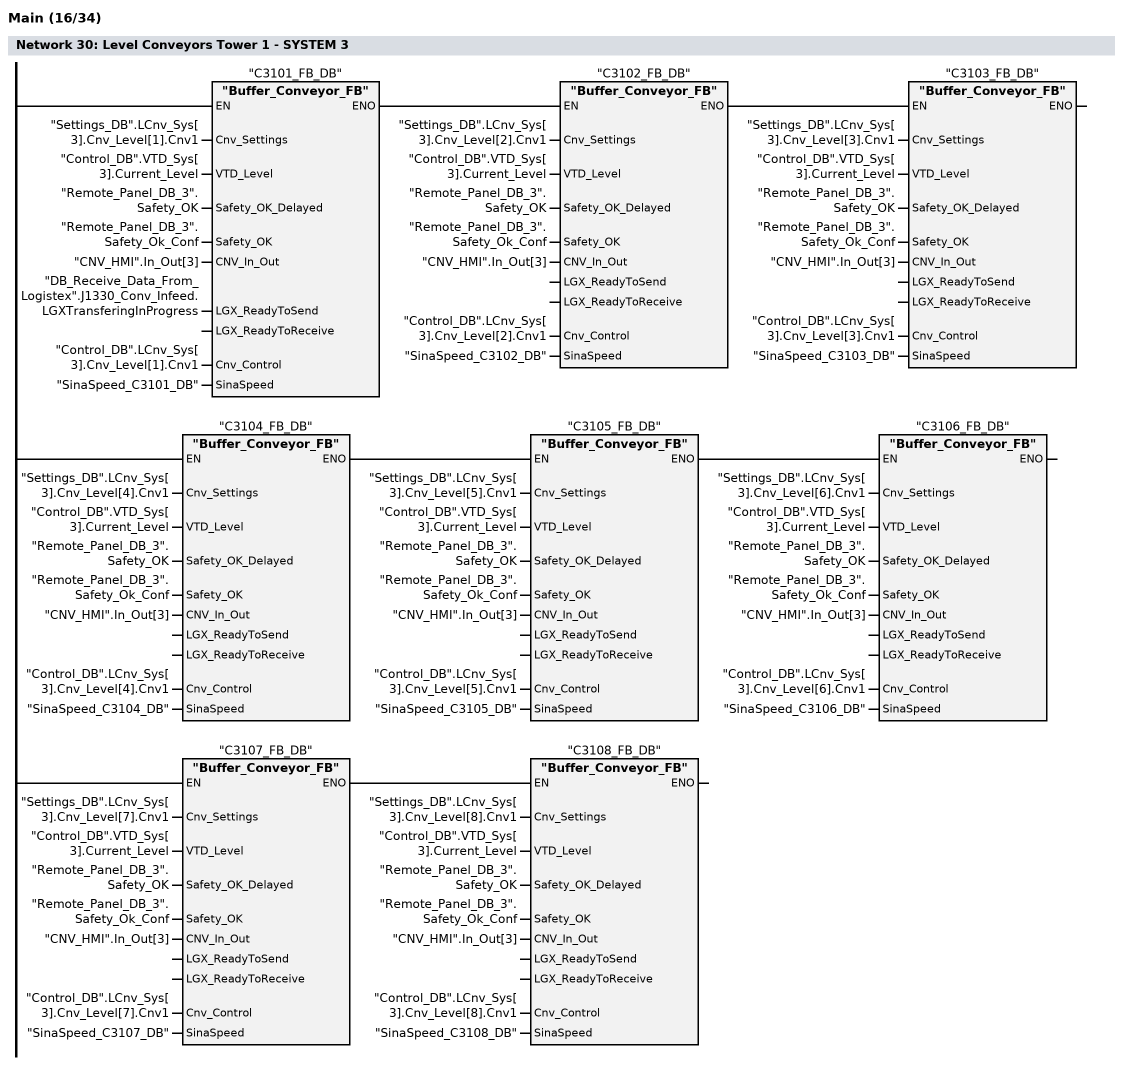
   RUNG wire#powerrail
      "C3101_FB_DB"(Cnv_Settings := "Settings_DB".LCnv_Sys[3].Cnv_Level[1].Cnv1, VTD_Level := "Control_DB".VTD_Sys[3].Current_Level, Safety_OK_Delayed := "Remote_Panel_DB_3".Safety_OK, Safety_OK := "Remote_Panel_DB_3".Safety_Ok_Conf, CNV_In_Out := "CNV_HMI".In_Out[3], LGX_ReadyToSend := "DB_Receive_Data_From_Logistex".J1330_Conv_Infeed.LGXTransferingInProgress, LGX_ReadyToReceive :=, Cnv_Control := "Control_DB".LCnv_Sys[3].Cnv_Level[1].Cnv1, SinaSpeed := "SinaSpeed_C3101_DB")
      "C3102_FB_DB"(Cnv_Settings := "Settings_DB".LCnv_Sys[3].Cnv_Level[2].Cnv1, VTD_Level := "Control_DB".VTD_Sys[3].Current_Level, Safety_OK_Delayed := "Remote_Panel_DB_3".Safety_OK, Safety_OK := "Remote_Panel_DB_3".Safety_Ok_Conf, CNV_In_Out := "CNV_HMI".In_Out[3], LGX_ReadyToSend :=, LGX_ReadyToReceive :=, Cnv_Control := "Control_DB".LCnv_Sys[3].Cnv_Level[2].Cnv1, SinaSpeed := "SinaSpeed_C3102_DB")
      "C3103_FB_DB"(Cnv_Settings := "Settings_DB".LCnv_Sys[3].Cnv_Level[3].Cnv1, VTD_Level := "Control_DB".VTD_Sys[3].Current_Level, Safety_OK_Delayed := "Remote_Panel_DB_3".Safety_OK, Safety_OK := "Remote_Panel_DB_3".Safety_Ok_Conf, CNV_In_Out := "CNV_HMI".In_Out[3], LGX_ReadyToSend :=, LGX_ReadyToReceive :=, Cnv_Control := "Control_DB".LCnv_Sys[3].Cnv_Level[3].Cnv1, SinaSpeed := "SinaSpeed_C3103_DB")
   END_RUNG
   RUNG wire#powerrail
      "C3104_FB_DB"(Cnv_Settings := "Settings_DB".LCnv_Sys[3].Cnv_Level[4].Cnv1, VTD_Level := "Control_DB".VTD_Sys[3].Current_Level, Safety_OK_Delayed := "Remote_Panel_DB_3".Safety_OK, Safety_OK := "Remote_Panel_DB_3".Safety_Ok_Conf, CNV_In_Out := "CNV_HMI".In_Out[3], LGX_ReadyToSend :=, LGX_ReadyToReceive :=, Cnv_Control := "Control_DB".LCnv_Sys[3].Cnv_Level[4].Cnv1, SinaSpeed := "SinaSpeed_C3104_DB")
      "C3105_FB_DB"(Cnv_Settings := "Settings_DB".LCnv_Sys[3].Cnv_Level[5].Cnv1, VTD_Level := "Control_DB".VTD_Sys[3].Current_Level, Safety_OK_Delayed := "Remote_Panel_DB_3".Safety_OK, Safety_OK := "Remote_Panel_DB_3".Safety_Ok_Conf, CNV_In_Out := "CNV_HMI".In_Out[3], LGX_ReadyToSend :=, LGX_ReadyToReceive :=, Cnv_Control := "Control_DB".LCnv_Sys[3].Cnv_Level[5].Cnv1, SinaSpeed := "SinaSpeed_C3105_DB")
      "C3106_FB_DB"(Cnv_Settings := "Settings_DB".LCnv_Sys[3].Cnv_Level[6].Cnv1, VTD_Level := "Control_DB".VTD_Sys[3].Current_Level, Safety_OK_Delayed := "Remote_Panel_DB_3".Safety_OK, Safety_OK := "Remote_Panel_DB_3".Safety_Ok_Conf, CNV_In_Out := "CNV_HMI".In_Out[3], LGX_ReadyToSend :=, LGX_ReadyToReceive :=, Cnv_Control := "Control_DB".LCnv_Sys[3].Cnv_Level[6].Cnv1, SinaSpeed := "SinaSpeed_C3106_DB")
   END_RUNG
   RUNG wire#powerrail
      "C3107_FB_DB"(Cnv_Settings := "Settings_DB".LCnv_Sys[3].Cnv_Level[7].Cnv1, VTD_Level := "Control_DB".VTD_Sys[3].Current_Level, Safety_OK_Delayed := "Remote_Panel_DB_3".Safety_OK, Safety_OK := "Remote_Panel_DB_3".Safety_Ok_Conf, CNV_In_Out := "CNV_HMI".In_Out[3], LGX_ReadyToSend :=, LGX_ReadyToReceive :=, Cnv_Control := "Control_DB".LCnv_Sys[3].Cnv_Level[7].Cnv1, SinaSpeed := "SinaSpeed_C3107_DB")
      "C3108_FB_DB"(Cnv_Settings := "Settings_DB".LCnv_Sys[3].Cnv_Level[8].Cnv1, VTD_Level := "Control_DB".VTD_Sys[3].Current_Level, Safety_OK_Delayed := "Remote_Panel_DB_3".Safety_OK, Safety_OK := "Remote_Panel_DB_3".Safety_Ok_Conf, CNV_In_Out := "CNV_HMI".In_Out[3], LGX_ReadyToSend :=, LGX_ReadyToReceive :=, Cnv_Control := "Control_DB".LCnv_Sys[3].Cnv_Level[8].Cnv1, SinaSpeed := "SinaSpeed_C3108_DB")
   END_RUNG
   // the same network as SCL:
   "C3101_FB_DB"(Cnv_Settings := "Settings_DB".LCnv_Sys[3].Cnv_Level[1].Cnv1,   // "Buffer_Conveyor_FB"
                 VTD_Level := "Control_DB".VTD_Sys[3].Current_Level,
                 Safety_OK_Delayed := "Remote_Panel_DB_3".Safety_OK,
                 Safety_OK := "Remote_Panel_DB_3".Safety_Ok_Conf,
                 CNV_In_Out := "CNV_HMI".In_Out[3],
                 LGX_ReadyToSend := "DB_Receive_Data_From_Logistex".J1330_Conv_Infeed.LGXTransferingInProgress,
                 Cnv_Control := "Control_DB".LCnv_Sys[3].Cnv_Level[1].Cnv1,
                 SinaSpeed := "SinaSpeed_C3101_DB",
                 ENO => #_w1);
   "C3102_FB_DB"(EN := #_w1,   // "Buffer_Conveyor_FB"
                 Cnv_Settings := "Settings_DB".LCnv_Sys[3].Cnv_Level[2].Cnv1,
                 VTD_Level := "Control_DB".VTD_Sys[3].Current_Level,
                 Safety_OK_Delayed := "Remote_Panel_DB_3".Safety_OK,
                 Safety_OK := "Remote_Panel_DB_3".Safety_Ok_Conf,
                 CNV_In_Out := "CNV_HMI".In_Out[3],
                 Cnv_Control := "Control_DB".LCnv_Sys[3].Cnv_Level[2].Cnv1,
                 SinaSpeed := "SinaSpeed_C3102_DB",
                 ENO => #_w2);
   IF #_w2 THEN
       "C3103_FB_DB"(Cnv_Settings := "Settings_DB".LCnv_Sys[3].Cnv_Level[3].Cnv1,   // "Buffer_Conveyor_FB"
                     VTD_Level := "Control_DB".VTD_Sys[3].Current_Level,
                     Safety_OK_Delayed := "Remote_Panel_DB_3".Safety_OK,
                     Safety_OK := "Remote_Panel_DB_3".Safety_Ok_Conf,
                     CNV_In_Out := "CNV_HMI".In_Out[3],
                     Cnv_Control := "Control_DB".LCnv_Sys[3].Cnv_Level[3].Cnv1,
                     SinaSpeed := "SinaSpeed_C3103_DB");
   END_IF;
   "C3104_FB_DB"(Cnv_Settings := "Settings_DB".LCnv_Sys[3].Cnv_Level[4].Cnv1,   // "Buffer_Conveyor_FB"
                 VTD_Level := "Control_DB".VTD_Sys[3].Current_Level,
                 Safety_OK_Delayed := "Remote_Panel_DB_3".Safety_OK,
                 Safety_OK := "Remote_Panel_DB_3".Safety_Ok_Conf,
                 CNV_In_Out := "CNV_HMI".In_Out[3],
                 Cnv_Control := "Control_DB".LCnv_Sys[3].Cnv_Level[4].Cnv1,
                 SinaSpeed := "SinaSpeed_C3104_DB",
                 ENO => #_w3);
   "C3105_FB_DB"(EN := #_w3,   // "Buffer_Conveyor_FB"
                 Cnv_Settings := "Settings_DB".LCnv_Sys[3].Cnv_Level[5].Cnv1,
                 VTD_Level := "Control_DB".VTD_Sys[3].Current_Level,
                 Safety_OK_Delayed := "Remote_Panel_DB_3".Safety_OK,
                 Safety_OK := "Remote_Panel_DB_3".Safety_Ok_Conf,
                 CNV_In_Out := "CNV_HMI".In_Out[3],
                 Cnv_Control := "Control_DB".LCnv_Sys[3].Cnv_Level[5].Cnv1,
                 SinaSpeed := "SinaSpeed_C3105_DB",
                 ENO => #_w4);
   IF #_w4 THEN
       "C3106_FB_DB"(Cnv_Settings := "Settings_DB".LCnv_Sys[3].Cnv_Level[6].Cnv1,   // "Buffer_Conveyor_FB"
                     VTD_Level := "Control_DB".VTD_Sys[3].Current_Level,
                     Safety_OK_Delayed := "Remote_Panel_DB_3".Safety_OK,
                     Safety_OK := "Remote_Panel_DB_3".Safety_Ok_Conf,
                     CNV_In_Out := "CNV_HMI".In_Out[3],
                     Cnv_Control := "Control_DB".LCnv_Sys[3].Cnv_Level[6].Cnv1,
                     SinaSpeed := "SinaSpeed_C3106_DB");
   END_IF;
   "C3107_FB_DB"(Cnv_Settings := "Settings_DB".LCnv_Sys[3].Cnv_Level[7].Cnv1,   // "Buffer_Conveyor_FB"
                 VTD_Level := "Control_DB".VTD_Sys[3].Current_Level,
                 Safety_OK_Delayed := "Remote_Panel_DB_3".Safety_OK,
                 Safety_OK := "Remote_Panel_DB_3".Safety_Ok_Conf,
                 CNV_In_Out := "CNV_HMI".In_Out[3],
                 Cnv_Control := "Control_DB".LCnv_Sys[3].Cnv_Level[7].Cnv1,
                 SinaSpeed := "SinaSpeed_C3107_DB",
                 ENO => #_w5);
   IF #_w5 THEN
       "C3108_FB_DB"(Cnv_Settings := "Settings_DB".LCnv_Sys[3].Cnv_Level[8].Cnv1,   // "Buffer_Conveyor_FB"
                     VTD_Level := "Control_DB".VTD_Sys[3].Current_Level,
                     Safety_OK_Delayed := "Remote_Panel_DB_3".Safety_OK,
                     Safety_OK := "Remote_Panel_DB_3".Safety_Ok_Conf,
                     CNV_In_Out := "CNV_HMI".In_Out[3],
                     Cnv_Control := "Control_DB".LCnv_Sys[3].Cnv_Level[8].Cnv1,
                     SinaSpeed := "SinaSpeed_C3108_DB");
   END_IF;
END_REGION

REGION Network 31: Level Conveyors Tower 2 - SYSTEM 3
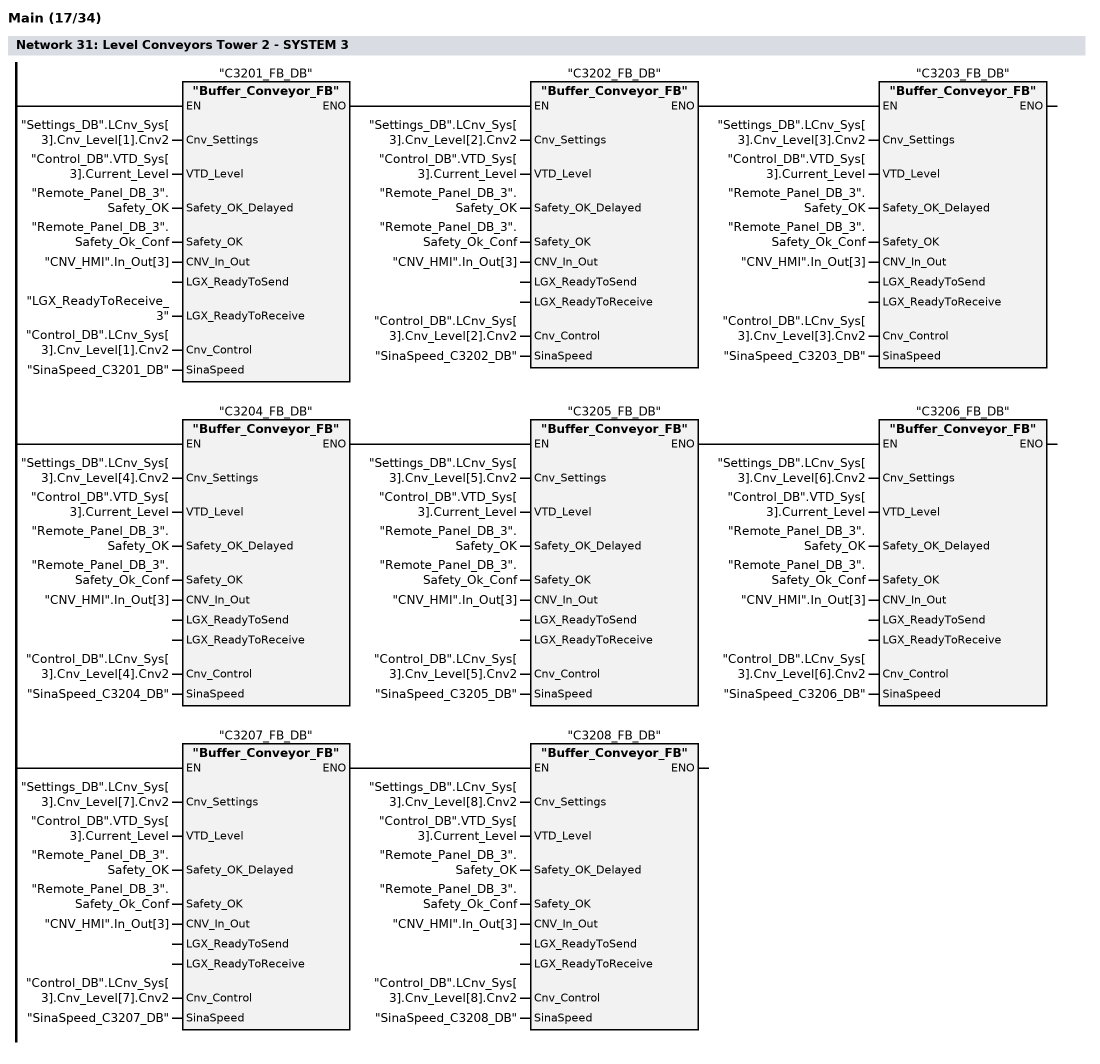
   RUNG wire#powerrail
      "C3201_FB_DB"(Cnv_Settings := "Settings_DB".LCnv_Sys[3].Cnv_Level[1].Cnv2, VTD_Level := "Control_DB".VTD_Sys[3].Current_Level, Safety_OK_Delayed := "Remote_Panel_DB_3".Safety_OK, Safety_OK := "Remote_Panel_DB_3".Safety_Ok_Conf, CNV_In_Out := "CNV_HMI".In_Out[3], LGX_ReadyToSend :=, LGX_ReadyToReceive := "LGX_ReadyToReceive_3", Cnv_Control := "Control_DB".LCnv_Sys[3].Cnv_Level[1].Cnv2, SinaSpeed := "SinaSpeed_C3201_DB")
      "C3202_FB_DB"(Cnv_Settings := "Settings_DB".LCnv_Sys[3].Cnv_Level[2].Cnv2, VTD_Level := "Control_DB".VTD_Sys[3].Current_Level, Safety_OK_Delayed := "Remote_Panel_DB_3".Safety_OK, Safety_OK := "Remote_Panel_DB_3".Safety_Ok_Conf, CNV_In_Out := "CNV_HMI".In_Out[3], LGX_ReadyToSend :=, LGX_ReadyToReceive :=, Cnv_Control := "Control_DB".LCnv_Sys[3].Cnv_Level[2].Cnv2, SinaSpeed := "SinaSpeed_C3202_DB")
      "C3203_FB_DB"(Cnv_Settings := "Settings_DB".LCnv_Sys[3].Cnv_Level[3].Cnv2, VTD_Level := "Control_DB".VTD_Sys[3].Current_Level, Safety_OK_Delayed := "Remote_Panel_DB_3".Safety_OK, Safety_OK := "Remote_Panel_DB_3".Safety_Ok_Conf, CNV_In_Out := "CNV_HMI".In_Out[3], LGX_ReadyToSend :=, LGX_ReadyToReceive :=, Cnv_Control := "Control_DB".LCnv_Sys[3].Cnv_Level[3].Cnv2, SinaSpeed := "SinaSpeed_C3203_DB")
   END_RUNG
   RUNG wire#powerrail
      "C3204_FB_DB"(Cnv_Settings := "Settings_DB".LCnv_Sys[3].Cnv_Level[4].Cnv2, VTD_Level := "Control_DB".VTD_Sys[3].Current_Level, Safety_OK_Delayed := "Remote_Panel_DB_3".Safety_OK, Safety_OK := "Remote_Panel_DB_3".Safety_Ok_Conf, CNV_In_Out := "CNV_HMI".In_Out[3], LGX_ReadyToSend :=, LGX_ReadyToReceive :=, Cnv_Control := "Control_DB".LCnv_Sys[3].Cnv_Level[4].Cnv2, SinaSpeed := "SinaSpeed_C3204_DB")
      "C3205_FB_DB"(Cnv_Settings := "Settings_DB".LCnv_Sys[3].Cnv_Level[5].Cnv2, VTD_Level := "Control_DB".VTD_Sys[3].Current_Level, Safety_OK_Delayed := "Remote_Panel_DB_3".Safety_OK, Safety_OK := "Remote_Panel_DB_3".Safety_Ok_Conf, CNV_In_Out := "CNV_HMI".In_Out[3], LGX_ReadyToSend :=, LGX_ReadyToReceive :=, Cnv_Control := "Control_DB".LCnv_Sys[3].Cnv_Level[5].Cnv2, SinaSpeed := "SinaSpeed_C3205_DB")
      "C3206_FB_DB"(Cnv_Settings := "Settings_DB".LCnv_Sys[3].Cnv_Level[6].Cnv2, VTD_Level := "Control_DB".VTD_Sys[3].Current_Level, Safety_OK_Delayed := "Remote_Panel_DB_3".Safety_OK, Safety_OK := "Remote_Panel_DB_3".Safety_Ok_Conf, CNV_In_Out := "CNV_HMI".In_Out[3], LGX_ReadyToSend :=, LGX_ReadyToReceive :=, Cnv_Control := "Control_DB".LCnv_Sys[3].Cnv_Level[6].Cnv2, SinaSpeed := "SinaSpeed_C3206_DB")
   END_RUNG
   RUNG wire#powerrail
      "C3207_FB_DB"(Cnv_Settings := "Settings_DB".LCnv_Sys[3].Cnv_Level[7].Cnv2, VTD_Level := "Control_DB".VTD_Sys[3].Current_Level, Safety_OK_Delayed := "Remote_Panel_DB_3".Safety_OK, Safety_OK := "Remote_Panel_DB_3".Safety_Ok_Conf, CNV_In_Out := "CNV_HMI".In_Out[3], LGX_ReadyToSend :=, LGX_ReadyToReceive :=, Cnv_Control := "Control_DB".LCnv_Sys[3].Cnv_Level[7].Cnv2, SinaSpeed := "SinaSpeed_C3207_DB")
      "C3208_FB_DB"(Cnv_Settings := "Settings_DB".LCnv_Sys[3].Cnv_Level[8].Cnv2, VTD_Level := "Control_DB".VTD_Sys[3].Current_Level, Safety_OK_Delayed := "Remote_Panel_DB_3".Safety_OK, Safety_OK := "Remote_Panel_DB_3".Safety_Ok_Conf, CNV_In_Out := "CNV_HMI".In_Out[3], LGX_ReadyToSend :=, LGX_ReadyToReceive :=, Cnv_Control := "Control_DB".LCnv_Sys[3].Cnv_Level[8].Cnv2, SinaSpeed := "SinaSpeed_C3208_DB")
   END_RUNG
   // the same network as SCL:
   "C3201_FB_DB"(Cnv_Settings := "Settings_DB".LCnv_Sys[3].Cnv_Level[1].Cnv2,   // "Buffer_Conveyor_FB"
                 VTD_Level := "Control_DB".VTD_Sys[3].Current_Level,
                 Safety_OK_Delayed := "Remote_Panel_DB_3".Safety_OK,
                 Safety_OK := "Remote_Panel_DB_3".Safety_Ok_Conf,
                 CNV_In_Out := "CNV_HMI".In_Out[3],
                 LGX_ReadyToReceive := "LGX_ReadyToReceive_3",
                 Cnv_Control := "Control_DB".LCnv_Sys[3].Cnv_Level[1].Cnv2,
                 SinaSpeed := "SinaSpeed_C3201_DB",
                 ENO => #_w1);
   "C3202_FB_DB"(EN := #_w1,   // "Buffer_Conveyor_FB"
                 Cnv_Settings := "Settings_DB".LCnv_Sys[3].Cnv_Level[2].Cnv2,
                 VTD_Level := "Control_DB".VTD_Sys[3].Current_Level,
                 Safety_OK_Delayed := "Remote_Panel_DB_3".Safety_OK,
                 Safety_OK := "Remote_Panel_DB_3".Safety_Ok_Conf,
                 CNV_In_Out := "CNV_HMI".In_Out[3],
                 Cnv_Control := "Control_DB".LCnv_Sys[3].Cnv_Level[2].Cnv2,
                 SinaSpeed := "SinaSpeed_C3202_DB",
                 ENO => #_w2);
   IF #_w2 THEN
       "C3203_FB_DB"(Cnv_Settings := "Settings_DB".LCnv_Sys[3].Cnv_Level[3].Cnv2,   // "Buffer_Conveyor_FB"
                     VTD_Level := "Control_DB".VTD_Sys[3].Current_Level,
                     Safety_OK_Delayed := "Remote_Panel_DB_3".Safety_OK,
                     Safety_OK := "Remote_Panel_DB_3".Safety_Ok_Conf,
                     CNV_In_Out := "CNV_HMI".In_Out[3],
                     Cnv_Control := "Control_DB".LCnv_Sys[3].Cnv_Level[3].Cnv2,
                     SinaSpeed := "SinaSpeed_C3203_DB");
   END_IF;
   "C3204_FB_DB"(Cnv_Settings := "Settings_DB".LCnv_Sys[3].Cnv_Level[4].Cnv2,   // "Buffer_Conveyor_FB"
                 VTD_Level := "Control_DB".VTD_Sys[3].Current_Level,
                 Safety_OK_Delayed := "Remote_Panel_DB_3".Safety_OK,
                 Safety_OK := "Remote_Panel_DB_3".Safety_Ok_Conf,
                 CNV_In_Out := "CNV_HMI".In_Out[3],
                 Cnv_Control := "Control_DB".LCnv_Sys[3].Cnv_Level[4].Cnv2,
                 SinaSpeed := "SinaSpeed_C3204_DB",
                 ENO => #_w3);
   "C3205_FB_DB"(EN := #_w3,   // "Buffer_Conveyor_FB"
                 Cnv_Settings := "Settings_DB".LCnv_Sys[3].Cnv_Level[5].Cnv2,
                 VTD_Level := "Control_DB".VTD_Sys[3].Current_Level,
                 Safety_OK_Delayed := "Remote_Panel_DB_3".Safety_OK,
                 Safety_OK := "Remote_Panel_DB_3".Safety_Ok_Conf,
                 CNV_In_Out := "CNV_HMI".In_Out[3],
                 Cnv_Control := "Control_DB".LCnv_Sys[3].Cnv_Level[5].Cnv2,
                 SinaSpeed := "SinaSpeed_C3205_DB",
                 ENO => #_w4);
   IF #_w4 THEN
       "C3206_FB_DB"(Cnv_Settings := "Settings_DB".LCnv_Sys[3].Cnv_Level[6].Cnv2,   // "Buffer_Conveyor_FB"
                     VTD_Level := "Control_DB".VTD_Sys[3].Current_Level,
                     Safety_OK_Delayed := "Remote_Panel_DB_3".Safety_OK,
                     Safety_OK := "Remote_Panel_DB_3".Safety_Ok_Conf,
                     CNV_In_Out := "CNV_HMI".In_Out[3],
                     Cnv_Control := "Control_DB".LCnv_Sys[3].Cnv_Level[6].Cnv2,
                     SinaSpeed := "SinaSpeed_C3206_DB");
   END_IF;
   "C3207_FB_DB"(Cnv_Settings := "Settings_DB".LCnv_Sys[3].Cnv_Level[7].Cnv2,   // "Buffer_Conveyor_FB"
                 VTD_Level := "Control_DB".VTD_Sys[3].Current_Level,
                 Safety_OK_Delayed := "Remote_Panel_DB_3".Safety_OK,
                 Safety_OK := "Remote_Panel_DB_3".Safety_Ok_Conf,
                 CNV_In_Out := "CNV_HMI".In_Out[3],
                 Cnv_Control := "Control_DB".LCnv_Sys[3].Cnv_Level[7].Cnv2,
                 SinaSpeed := "SinaSpeed_C3207_DB",
                 ENO => #_w5);
   IF #_w5 THEN
       "C3208_FB_DB"(Cnv_Settings := "Settings_DB".LCnv_Sys[3].Cnv_Level[8].Cnv2,   // "Buffer_Conveyor_FB"
                     VTD_Level := "Control_DB".VTD_Sys[3].Current_Level,
                     Safety_OK_Delayed := "Remote_Panel_DB_3".Safety_OK,
                     Safety_OK := "Remote_Panel_DB_3".Safety_Ok_Conf,
                     CNV_In_Out := "CNV_HMI".In_Out[3],
                     Cnv_Control := "Control_DB".LCnv_Sys[3].Cnv_Level[8].Cnv2,
                     SinaSpeed := "SinaSpeed_C3208_DB");
   END_IF;
END_REGION

REGION Network 32: SAFETY STOPPERS Tower 1 - SYSTEM 3
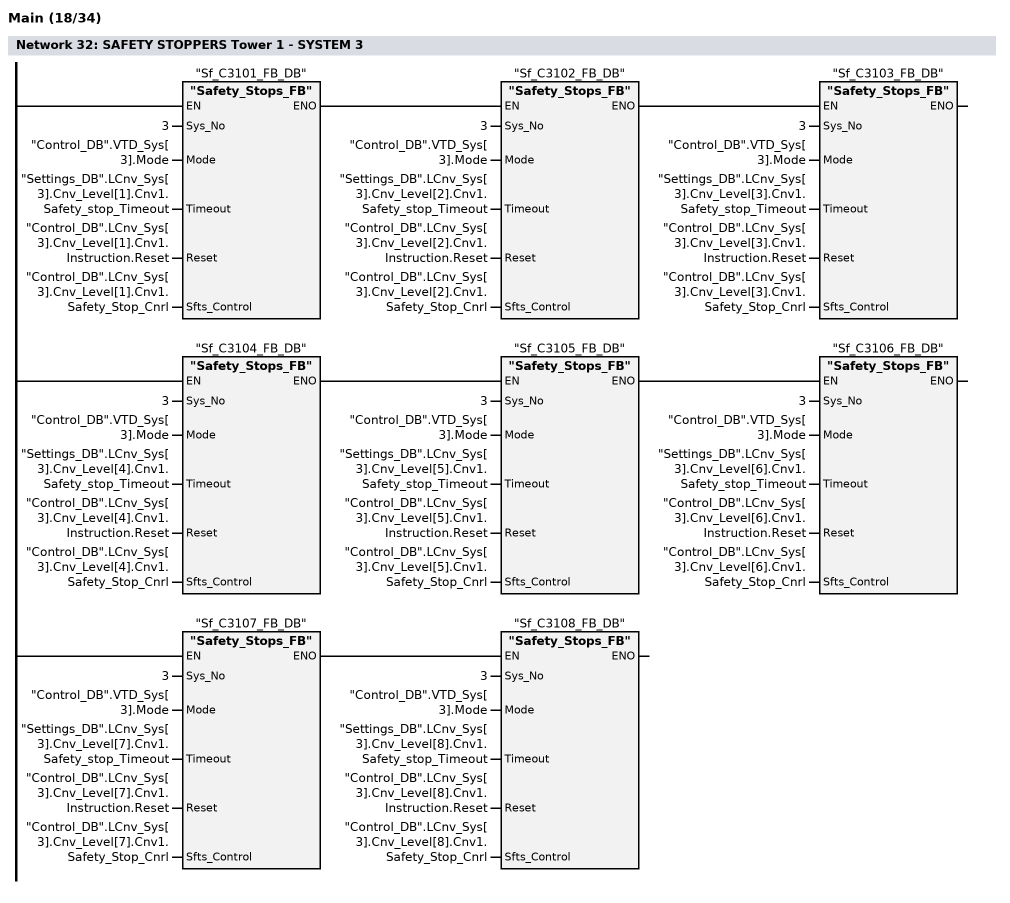
   RUNG wire#powerrail
      "Sf_C3101_FB_DB"(Sys_No := 3, Mode := "Control_DB".VTD_Sys[3].Mode, Timeout := "Settings_DB".LCnv_Sys[3].Cnv_Level[1].Cnv1.Safety_stop_Timeout, Reset := "Control_DB".LCnv_Sys[3].Cnv_Level[1].Cnv1.Instruction.Reset, Sfts_Control := "Control_DB".LCnv_Sys[3].Cnv_Level[1].Cnv1.Safety_Stop_Cnrl)
      "Sf_C3102_FB_DB"(Sys_No := 3, Mode := "Control_DB".VTD_Sys[3].Mode, Timeout := "Settings_DB".LCnv_Sys[3].Cnv_Level[2].Cnv1.Safety_stop_Timeout, Reset := "Control_DB".LCnv_Sys[3].Cnv_Level[2].Cnv1.Instruction.Reset, Sfts_Control := "Control_DB".LCnv_Sys[3].Cnv_Level[2].Cnv1.Safety_Stop_Cnrl)
      "Sf_C3103_FB_DB"(Sys_No := 3, Mode := "Control_DB".VTD_Sys[3].Mode, Timeout := "Settings_DB".LCnv_Sys[3].Cnv_Level[3].Cnv1.Safety_stop_Timeout, Reset := "Control_DB".LCnv_Sys[3].Cnv_Level[3].Cnv1.Instruction.Reset, Sfts_Control := "Control_DB".LCnv_Sys[3].Cnv_Level[3].Cnv1.Safety_Stop_Cnrl)
   END_RUNG
   RUNG wire#powerrail
      "Sf_C3104_FB_DB"(Sys_No := 3, Mode := "Control_DB".VTD_Sys[3].Mode, Timeout := "Settings_DB".LCnv_Sys[3].Cnv_Level[4].Cnv1.Safety_stop_Timeout, Reset := "Control_DB".LCnv_Sys[3].Cnv_Level[4].Cnv1.Instruction.Reset, Sfts_Control := "Control_DB".LCnv_Sys[3].Cnv_Level[4].Cnv1.Safety_Stop_Cnrl)
      "Sf_C3105_FB_DB"(Sys_No := 3, Mode := "Control_DB".VTD_Sys[3].Mode, Timeout := "Settings_DB".LCnv_Sys[3].Cnv_Level[5].Cnv1.Safety_stop_Timeout, Reset := "Control_DB".LCnv_Sys[3].Cnv_Level[5].Cnv1.Instruction.Reset, Sfts_Control := "Control_DB".LCnv_Sys[3].Cnv_Level[5].Cnv1.Safety_Stop_Cnrl)
      "Sf_C3106_FB_DB"(Sys_No := 3, Mode := "Control_DB".VTD_Sys[3].Mode, Timeout := "Settings_DB".LCnv_Sys[3].Cnv_Level[6].Cnv1.Safety_stop_Timeout, Reset := "Control_DB".LCnv_Sys[3].Cnv_Level[6].Cnv1.Instruction.Reset, Sfts_Control := "Control_DB".LCnv_Sys[3].Cnv_Level[6].Cnv1.Safety_Stop_Cnrl)
   END_RUNG
   RUNG wire#powerrail
      "Sf_C3107_FB_DB"(Sys_No := 3, Mode := "Control_DB".VTD_Sys[3].Mode, Timeout := "Settings_DB".LCnv_Sys[3].Cnv_Level[7].Cnv1.Safety_stop_Timeout, Reset := "Control_DB".LCnv_Sys[3].Cnv_Level[7].Cnv1.Instruction.Reset, Sfts_Control := "Control_DB".LCnv_Sys[3].Cnv_Level[7].Cnv1.Safety_Stop_Cnrl)
      "Sf_C3108_FB_DB"(Sys_No := 3, Mode := "Control_DB".VTD_Sys[3].Mode, Timeout := "Settings_DB".LCnv_Sys[3].Cnv_Level[8].Cnv1.Safety_stop_Timeout, Reset := "Control_DB".LCnv_Sys[3].Cnv_Level[8].Cnv1.Instruction.Reset, Sfts_Control := "Control_DB".LCnv_Sys[3].Cnv_Level[8].Cnv1.Safety_Stop_Cnrl)
   END_RUNG
   // the same network as SCL:
   "Sf_C3101_FB_DB"(Sys_No := 3,   // "Safety_Stops_FB"
                    Mode := "Control_DB".VTD_Sys[3].Mode,
                    Timeout := "Settings_DB".LCnv_Sys[3].Cnv_Level[1].Cnv1.Safety_stop_Timeout,
                    Reset := "Control_DB".LCnv_Sys[3].Cnv_Level[1].Cnv1.Instruction.Reset,
                    Sfts_Control := "Control_DB".LCnv_Sys[3].Cnv_Level[1].Cnv1.Safety_Stop_Cnrl,
                    ENO => #_w1);
   "Sf_C3102_FB_DB"(EN := #_w1,   // "Safety_Stops_FB"
                    Sys_No := 3,
                    Mode := "Control_DB".VTD_Sys[3].Mode,
                    Timeout := "Settings_DB".LCnv_Sys[3].Cnv_Level[2].Cnv1.Safety_stop_Timeout,
                    Reset := "Control_DB".LCnv_Sys[3].Cnv_Level[2].Cnv1.Instruction.Reset,
                    Sfts_Control := "Control_DB".LCnv_Sys[3].Cnv_Level[2].Cnv1.Safety_Stop_Cnrl,
                    ENO => #_w2);
   IF #_w2 THEN
       "Sf_C3103_FB_DB"(Sys_No := 3,   // "Safety_Stops_FB"
                        Mode := "Control_DB".VTD_Sys[3].Mode,
                        Timeout := "Settings_DB".LCnv_Sys[3].Cnv_Level[3].Cnv1.Safety_stop_Timeout,
                        Reset := "Control_DB".LCnv_Sys[3].Cnv_Level[3].Cnv1.Instruction.Reset,
                        Sfts_Control := "Control_DB".LCnv_Sys[3].Cnv_Level[3].Cnv1.Safety_Stop_Cnrl);
   END_IF;
   "Sf_C3104_FB_DB"(Sys_No := 3,   // "Safety_Stops_FB"
                    Mode := "Control_DB".VTD_Sys[3].Mode,
                    Timeout := "Settings_DB".LCnv_Sys[3].Cnv_Level[4].Cnv1.Safety_stop_Timeout,
                    Reset := "Control_DB".LCnv_Sys[3].Cnv_Level[4].Cnv1.Instruction.Reset,
                    Sfts_Control := "Control_DB".LCnv_Sys[3].Cnv_Level[4].Cnv1.Safety_Stop_Cnrl,
                    ENO => #_w3);
   "Sf_C3105_FB_DB"(EN := #_w3,   // "Safety_Stops_FB"
                    Sys_No := 3,
                    Mode := "Control_DB".VTD_Sys[3].Mode,
                    Timeout := "Settings_DB".LCnv_Sys[3].Cnv_Level[5].Cnv1.Safety_stop_Timeout,
                    Reset := "Control_DB".LCnv_Sys[3].Cnv_Level[5].Cnv1.Instruction.Reset,
                    Sfts_Control := "Control_DB".LCnv_Sys[3].Cnv_Level[5].Cnv1.Safety_Stop_Cnrl,
                    ENO => #_w4);
   IF #_w4 THEN
       "Sf_C3106_FB_DB"(Sys_No := 3,   // "Safety_Stops_FB"
                        Mode := "Control_DB".VTD_Sys[3].Mode,
                        Timeout := "Settings_DB".LCnv_Sys[3].Cnv_Level[6].Cnv1.Safety_stop_Timeout,
                        Reset := "Control_DB".LCnv_Sys[3].Cnv_Level[6].Cnv1.Instruction.Reset,
                        Sfts_Control := "Control_DB".LCnv_Sys[3].Cnv_Level[6].Cnv1.Safety_Stop_Cnrl);
   END_IF;
   "Sf_C3107_FB_DB"(Sys_No := 3,   // "Safety_Stops_FB"
                    Mode := "Control_DB".VTD_Sys[3].Mode,
                    Timeout := "Settings_DB".LCnv_Sys[3].Cnv_Level[7].Cnv1.Safety_stop_Timeout,
                    Reset := "Control_DB".LCnv_Sys[3].Cnv_Level[7].Cnv1.Instruction.Reset,
                    Sfts_Control := "Control_DB".LCnv_Sys[3].Cnv_Level[7].Cnv1.Safety_Stop_Cnrl,
                    ENO => #_w5);
   IF #_w5 THEN
       "Sf_C3108_FB_DB"(Sys_No := 3,   // "Safety_Stops_FB"
                        Mode := "Control_DB".VTD_Sys[3].Mode,
                        Timeout := "Settings_DB".LCnv_Sys[3].Cnv_Level[8].Cnv1.Safety_stop_Timeout,
                        Reset := "Control_DB".LCnv_Sys[3].Cnv_Level[8].Cnv1.Instruction.Reset,
                        Sfts_Control := "Control_DB".LCnv_Sys[3].Cnv_Level[8].Cnv1.Safety_Stop_Cnrl);
   END_IF;
END_REGION

REGION Network 33: SAFETY STOPPERS Tower 2 - SYSTEM 3
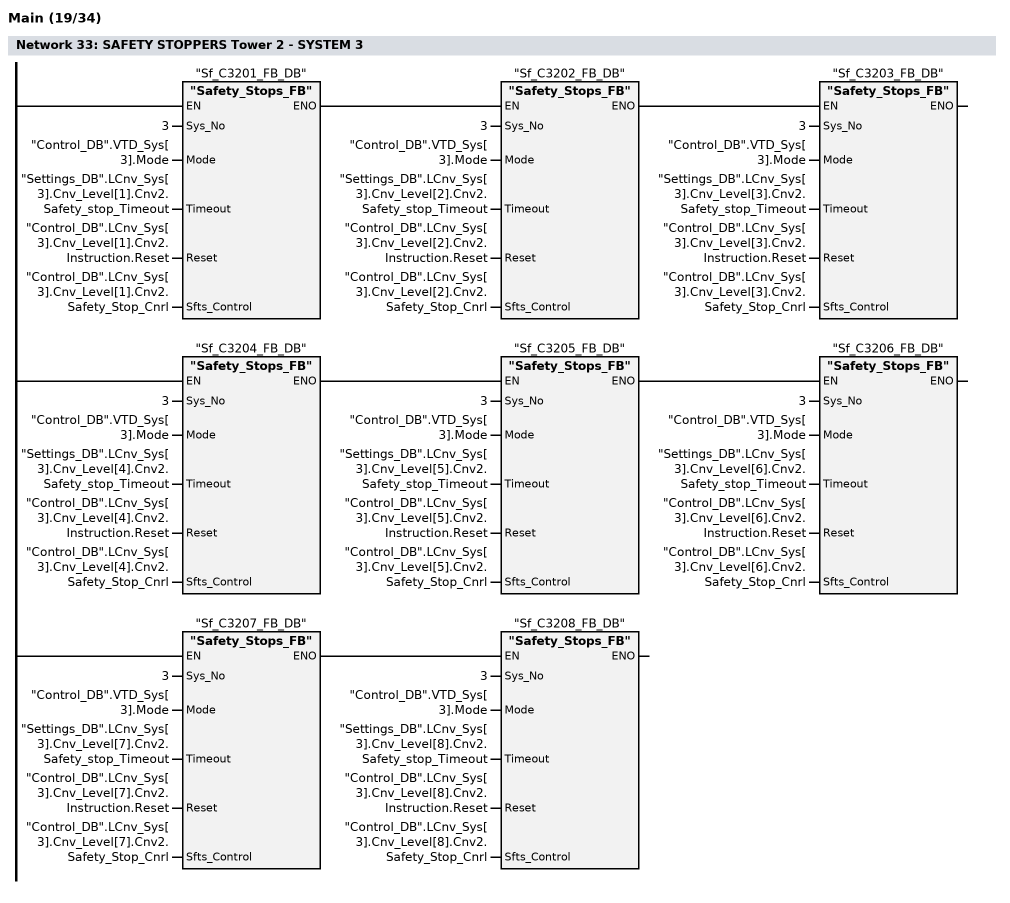
   RUNG wire#powerrail
      "Sf_C3201_FB_DB"(Sys_No := 3, Mode := "Control_DB".VTD_Sys[3].Mode, Timeout := "Settings_DB".LCnv_Sys[3].Cnv_Level[1].Cnv2.Safety_stop_Timeout, Reset := "Control_DB".LCnv_Sys[3].Cnv_Level[1].Cnv2.Instruction.Reset, Sfts_Control := "Control_DB".LCnv_Sys[3].Cnv_Level[1].Cnv2.Safety_Stop_Cnrl)
      "Sf_C3202_FB_DB"(Sys_No := 3, Mode := "Control_DB".VTD_Sys[3].Mode, Timeout := "Settings_DB".LCnv_Sys[3].Cnv_Level[2].Cnv2.Safety_stop_Timeout, Reset := "Control_DB".LCnv_Sys[3].Cnv_Level[2].Cnv2.Instruction.Reset, Sfts_Control := "Control_DB".LCnv_Sys[3].Cnv_Level[2].Cnv2.Safety_Stop_Cnrl)
      "Sf_C3203_FB_DB"(Sys_No := 3, Mode := "Control_DB".VTD_Sys[3].Mode, Timeout := "Settings_DB".LCnv_Sys[3].Cnv_Level[3].Cnv2.Safety_stop_Timeout, Reset := "Control_DB".LCnv_Sys[3].Cnv_Level[3].Cnv2.Instruction.Reset, Sfts_Control := "Control_DB".LCnv_Sys[3].Cnv_Level[3].Cnv2.Safety_Stop_Cnrl)
   END_RUNG
   RUNG wire#powerrail
      "Sf_C3204_FB_DB"(Sys_No := 3, Mode := "Control_DB".VTD_Sys[3].Mode, Timeout := "Settings_DB".LCnv_Sys[3].Cnv_Level[4].Cnv2.Safety_stop_Timeout, Reset := "Control_DB".LCnv_Sys[3].Cnv_Level[4].Cnv2.Instruction.Reset, Sfts_Control := "Control_DB".LCnv_Sys[3].Cnv_Level[4].Cnv2.Safety_Stop_Cnrl)
      "Sf_C3205_FB_DB"(Sys_No := 3, Mode := "Control_DB".VTD_Sys[3].Mode, Timeout := "Settings_DB".LCnv_Sys[3].Cnv_Level[5].Cnv2.Safety_stop_Timeout, Reset := "Control_DB".LCnv_Sys[3].Cnv_Level[5].Cnv2.Instruction.Reset, Sfts_Control := "Control_DB".LCnv_Sys[3].Cnv_Level[5].Cnv2.Safety_Stop_Cnrl)
      "Sf_C3206_FB_DB"(Sys_No := 3, Mode := "Control_DB".VTD_Sys[3].Mode, Timeout := "Settings_DB".LCnv_Sys[3].Cnv_Level[6].Cnv2.Safety_stop_Timeout, Reset := "Control_DB".LCnv_Sys[3].Cnv_Level[6].Cnv2.Instruction.Reset, Sfts_Control := "Control_DB".LCnv_Sys[3].Cnv_Level[6].Cnv2.Safety_Stop_Cnrl)
   END_RUNG
   RUNG wire#powerrail
      "Sf_C3207_FB_DB"(Sys_No := 3, Mode := "Control_DB".VTD_Sys[3].Mode, Timeout := "Settings_DB".LCnv_Sys[3].Cnv_Level[7].Cnv2.Safety_stop_Timeout, Reset := "Control_DB".LCnv_Sys[3].Cnv_Level[7].Cnv2.Instruction.Reset, Sfts_Control := "Control_DB".LCnv_Sys[3].Cnv_Level[7].Cnv2.Safety_Stop_Cnrl)
      "Sf_C3208_FB_DB"(Sys_No := 3, Mode := "Control_DB".VTD_Sys[3].Mode, Timeout := "Settings_DB".LCnv_Sys[3].Cnv_Level[8].Cnv2.Safety_stop_Timeout, Reset := "Control_DB".LCnv_Sys[3].Cnv_Level[8].Cnv2.Instruction.Reset, Sfts_Control := "Control_DB".LCnv_Sys[3].Cnv_Level[8].Cnv2.Safety_Stop_Cnrl)
   END_RUNG
   // the same network as SCL:
   "Sf_C3201_FB_DB"(Sys_No := 3,   // "Safety_Stops_FB"
                    Mode := "Control_DB".VTD_Sys[3].Mode,
                    Timeout := "Settings_DB".LCnv_Sys[3].Cnv_Level[1].Cnv2.Safety_stop_Timeout,
                    Reset := "Control_DB".LCnv_Sys[3].Cnv_Level[1].Cnv2.Instruction.Reset,
                    Sfts_Control := "Control_DB".LCnv_Sys[3].Cnv_Level[1].Cnv2.Safety_Stop_Cnrl,
                    ENO => #_w1);
   "Sf_C3202_FB_DB"(EN := #_w1,   // "Safety_Stops_FB"
                    Sys_No := 3,
                    Mode := "Control_DB".VTD_Sys[3].Mode,
                    Timeout := "Settings_DB".LCnv_Sys[3].Cnv_Level[2].Cnv2.Safety_stop_Timeout,
                    Reset := "Control_DB".LCnv_Sys[3].Cnv_Level[2].Cnv2.Instruction.Reset,
                    Sfts_Control := "Control_DB".LCnv_Sys[3].Cnv_Level[2].Cnv2.Safety_Stop_Cnrl,
                    ENO => #_w2);
   IF #_w2 THEN
       "Sf_C3203_FB_DB"(Sys_No := 3,   // "Safety_Stops_FB"
                        Mode := "Control_DB".VTD_Sys[3].Mode,
                        Timeout := "Settings_DB".LCnv_Sys[3].Cnv_Level[3].Cnv2.Safety_stop_Timeout,
                        Reset := "Control_DB".LCnv_Sys[3].Cnv_Level[3].Cnv2.Instruction.Reset,
                        Sfts_Control := "Control_DB".LCnv_Sys[3].Cnv_Level[3].Cnv2.Safety_Stop_Cnrl);
   END_IF;
   "Sf_C3204_FB_DB"(Sys_No := 3,   // "Safety_Stops_FB"
                    Mode := "Control_DB".VTD_Sys[3].Mode,
                    Timeout := "Settings_DB".LCnv_Sys[3].Cnv_Level[4].Cnv2.Safety_stop_Timeout,
                    Reset := "Control_DB".LCnv_Sys[3].Cnv_Level[4].Cnv2.Instruction.Reset,
                    Sfts_Control := "Control_DB".LCnv_Sys[3].Cnv_Level[4].Cnv2.Safety_Stop_Cnrl,
                    ENO => #_w3);
   "Sf_C3205_FB_DB"(EN := #_w3,   // "Safety_Stops_FB"
                    Sys_No := 3,
                    Mode := "Control_DB".VTD_Sys[3].Mode,
                    Timeout := "Settings_DB".LCnv_Sys[3].Cnv_Level[5].Cnv2.Safety_stop_Timeout,
                    Reset := "Control_DB".LCnv_Sys[3].Cnv_Level[5].Cnv2.Instruction.Reset,
                    Sfts_Control := "Control_DB".LCnv_Sys[3].Cnv_Level[5].Cnv2.Safety_Stop_Cnrl,
                    ENO => #_w4);
   IF #_w4 THEN
       "Sf_C3206_FB_DB"(Sys_No := 3,   // "Safety_Stops_FB"
                        Mode := "Control_DB".VTD_Sys[3].Mode,
                        Timeout := "Settings_DB".LCnv_Sys[3].Cnv_Level[6].Cnv2.Safety_stop_Timeout,
                        Reset := "Control_DB".LCnv_Sys[3].Cnv_Level[6].Cnv2.Instruction.Reset,
                        Sfts_Control := "Control_DB".LCnv_Sys[3].Cnv_Level[6].Cnv2.Safety_Stop_Cnrl);
   END_IF;
   "Sf_C3207_FB_DB"(Sys_No := 3,   // "Safety_Stops_FB"
                    Mode := "Control_DB".VTD_Sys[3].Mode,
                    Timeout := "Settings_DB".LCnv_Sys[3].Cnv_Level[7].Cnv2.Safety_stop_Timeout,
                    Reset := "Control_DB".LCnv_Sys[3].Cnv_Level[7].Cnv2.Instruction.Reset,
                    Sfts_Control := "Control_DB".LCnv_Sys[3].Cnv_Level[7].Cnv2.Safety_Stop_Cnrl,
                    ENO => #_w5);
   IF #_w5 THEN
       "Sf_C3208_FB_DB"(Sys_No := 3,   // "Safety_Stops_FB"
                        Mode := "Control_DB".VTD_Sys[3].Mode,
                        Timeout := "Settings_DB".LCnv_Sys[3].Cnv_Level[8].Cnv2.Safety_stop_Timeout,
                        Reset := "Control_DB".LCnv_Sys[3].Cnv_Level[8].Cnv2.Instruction.Reset,
                        Sfts_Control := "Control_DB".LCnv_Sys[3].Cnv_Level[8].Cnv2.Safety_Stop_Cnrl);
   END_IF;
END_REGION

REGION Network 34: SYSTEM 4
END_REGION

REGION Network 35: Level Conveyors Tower 1 - SYSTEM 4
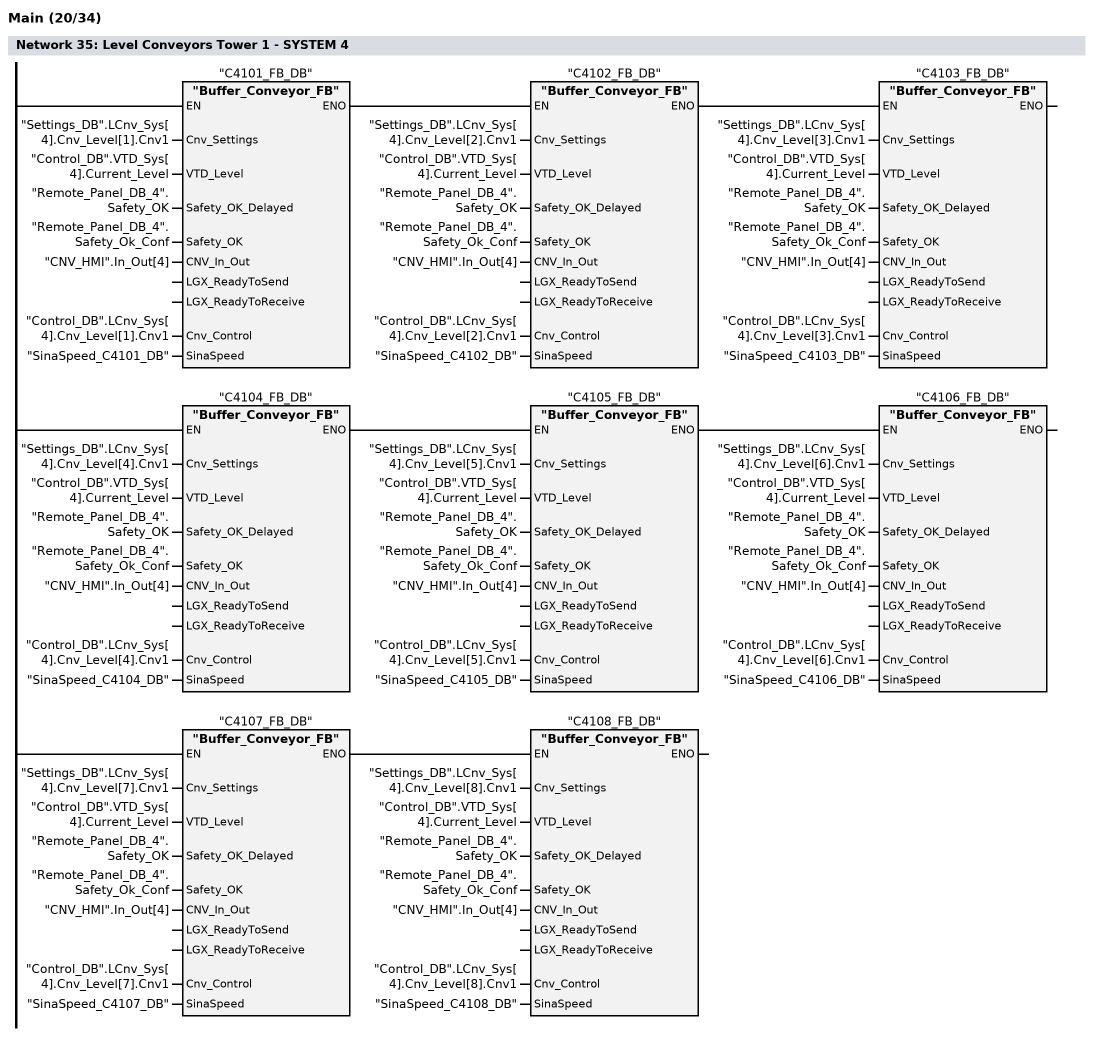
   RUNG wire#powerrail
      "C4101_FB_DB"(Cnv_Settings := "Settings_DB".LCnv_Sys[4].Cnv_Level[1].Cnv1, VTD_Level := "Control_DB".VTD_Sys[4].Current_Level, Safety_OK_Delayed := "Remote_Panel_DB_4".Safety_OK, Safety_OK := "Remote_Panel_DB_4".Safety_Ok_Conf, CNV_In_Out := "CNV_HMI".In_Out[4], LGX_ReadyToSend :=, LGX_ReadyToReceive :=, Cnv_Control := "Control_DB".LCnv_Sys[4].Cnv_Level[1].Cnv1, SinaSpeed := "SinaSpeed_C4101_DB")
      "C4102_FB_DB"(Cnv_Settings := "Settings_DB".LCnv_Sys[4].Cnv_Level[2].Cnv1, VTD_Level := "Control_DB".VTD_Sys[4].Current_Level, Safety_OK_Delayed := "Remote_Panel_DB_4".Safety_OK, Safety_OK := "Remote_Panel_DB_4".Safety_Ok_Conf, CNV_In_Out := "CNV_HMI".In_Out[4], LGX_ReadyToSend :=, LGX_ReadyToReceive :=, Cnv_Control := "Control_DB".LCnv_Sys[4].Cnv_Level[2].Cnv1, SinaSpeed := "SinaSpeed_C4102_DB")
      "C4103_FB_DB"(Cnv_Settings := "Settings_DB".LCnv_Sys[4].Cnv_Level[3].Cnv1, VTD_Level := "Control_DB".VTD_Sys[4].Current_Level, Safety_OK_Delayed := "Remote_Panel_DB_4".Safety_OK, Safety_OK := "Remote_Panel_DB_4".Safety_Ok_Conf, CNV_In_Out := "CNV_HMI".In_Out[4], LGX_ReadyToSend :=, LGX_ReadyToReceive :=, Cnv_Control := "Control_DB".LCnv_Sys[4].Cnv_Level[3].Cnv1, SinaSpeed := "SinaSpeed_C4103_DB")
   END_RUNG
   RUNG wire#powerrail
      "C4104_FB_DB"(Cnv_Settings := "Settings_DB".LCnv_Sys[4].Cnv_Level[4].Cnv1, VTD_Level := "Control_DB".VTD_Sys[4].Current_Level, Safety_OK_Delayed := "Remote_Panel_DB_4".Safety_OK, Safety_OK := "Remote_Panel_DB_4".Safety_Ok_Conf, CNV_In_Out := "CNV_HMI".In_Out[4], LGX_ReadyToSend :=, LGX_ReadyToReceive :=, Cnv_Control := "Control_DB".LCnv_Sys[4].Cnv_Level[4].Cnv1, SinaSpeed := "SinaSpeed_C4104_DB")
      "C4105_FB_DB"(Cnv_Settings := "Settings_DB".LCnv_Sys[4].Cnv_Level[5].Cnv1, VTD_Level := "Control_DB".VTD_Sys[4].Current_Level, Safety_OK_Delayed := "Remote_Panel_DB_4".Safety_OK, Safety_OK := "Remote_Panel_DB_4".Safety_Ok_Conf, CNV_In_Out := "CNV_HMI".In_Out[4], LGX_ReadyToSend :=, LGX_ReadyToReceive :=, Cnv_Control := "Control_DB".LCnv_Sys[4].Cnv_Level[5].Cnv1, SinaSpeed := "SinaSpeed_C4105_DB")
      "C4106_FB_DB"(Cnv_Settings := "Settings_DB".LCnv_Sys[4].Cnv_Level[6].Cnv1, VTD_Level := "Control_DB".VTD_Sys[4].Current_Level, Safety_OK_Delayed := "Remote_Panel_DB_4".Safety_OK, Safety_OK := "Remote_Panel_DB_4".Safety_Ok_Conf, CNV_In_Out := "CNV_HMI".In_Out[4], LGX_ReadyToSend :=, LGX_ReadyToReceive :=, Cnv_Control := "Control_DB".LCnv_Sys[4].Cnv_Level[6].Cnv1, SinaSpeed := "SinaSpeed_C4106_DB")
   END_RUNG
   RUNG wire#powerrail
      "C4107_FB_DB"(Cnv_Settings := "Settings_DB".LCnv_Sys[4].Cnv_Level[7].Cnv1, VTD_Level := "Control_DB".VTD_Sys[4].Current_Level, Safety_OK_Delayed := "Remote_Panel_DB_4".Safety_OK, Safety_OK := "Remote_Panel_DB_4".Safety_Ok_Conf, CNV_In_Out := "CNV_HMI".In_Out[4], LGX_ReadyToSend :=, LGX_ReadyToReceive :=, Cnv_Control := "Control_DB".LCnv_Sys[4].Cnv_Level[7].Cnv1, SinaSpeed := "SinaSpeed_C4107_DB")
      "C4108_FB_DB"(Cnv_Settings := "Settings_DB".LCnv_Sys[4].Cnv_Level[8].Cnv1, VTD_Level := "Control_DB".VTD_Sys[4].Current_Level, Safety_OK_Delayed := "Remote_Panel_DB_4".Safety_OK, Safety_OK := "Remote_Panel_DB_4".Safety_Ok_Conf, CNV_In_Out := "CNV_HMI".In_Out[4], LGX_ReadyToSend :=, LGX_ReadyToReceive :=, Cnv_Control := "Control_DB".LCnv_Sys[4].Cnv_Level[8].Cnv1, SinaSpeed := "SinaSpeed_C4108_DB")
   END_RUNG
   // the same network as SCL:
   "C4101_FB_DB"(Cnv_Settings := "Settings_DB".LCnv_Sys[4].Cnv_Level[1].Cnv1,   // "Buffer_Conveyor_FB"
                 VTD_Level := "Control_DB".VTD_Sys[4].Current_Level,
                 Safety_OK_Delayed := "Remote_Panel_DB_4".Safety_OK,
                 Safety_OK := "Remote_Panel_DB_4".Safety_Ok_Conf,
                 CNV_In_Out := "CNV_HMI".In_Out[4],
                 Cnv_Control := "Control_DB".LCnv_Sys[4].Cnv_Level[1].Cnv1,
                 SinaSpeed := "SinaSpeed_C4101_DB",
                 ENO => #_w1);
   "C4102_FB_DB"(EN := #_w1,   // "Buffer_Conveyor_FB"
                 Cnv_Settings := "Settings_DB".LCnv_Sys[4].Cnv_Level[2].Cnv1,
                 VTD_Level := "Control_DB".VTD_Sys[4].Current_Level,
                 Safety_OK_Delayed := "Remote_Panel_DB_4".Safety_OK,
                 Safety_OK := "Remote_Panel_DB_4".Safety_Ok_Conf,
                 CNV_In_Out := "CNV_HMI".In_Out[4],
                 Cnv_Control := "Control_DB".LCnv_Sys[4].Cnv_Level[2].Cnv1,
                 SinaSpeed := "SinaSpeed_C4102_DB",
                 ENO => #_w2);
   IF #_w2 THEN
       "C4103_FB_DB"(Cnv_Settings := "Settings_DB".LCnv_Sys[4].Cnv_Level[3].Cnv1,   // "Buffer_Conveyor_FB"
                     VTD_Level := "Control_DB".VTD_Sys[4].Current_Level,
                     Safety_OK_Delayed := "Remote_Panel_DB_4".Safety_OK,
                     Safety_OK := "Remote_Panel_DB_4".Safety_Ok_Conf,
                     CNV_In_Out := "CNV_HMI".In_Out[4],
                     Cnv_Control := "Control_DB".LCnv_Sys[4].Cnv_Level[3].Cnv1,
                     SinaSpeed := "SinaSpeed_C4103_DB");
   END_IF;
   "C4104_FB_DB"(Cnv_Settings := "Settings_DB".LCnv_Sys[4].Cnv_Level[4].Cnv1,   // "Buffer_Conveyor_FB"
                 VTD_Level := "Control_DB".VTD_Sys[4].Current_Level,
                 Safety_OK_Delayed := "Remote_Panel_DB_4".Safety_OK,
                 Safety_OK := "Remote_Panel_DB_4".Safety_Ok_Conf,
                 CNV_In_Out := "CNV_HMI".In_Out[4],
                 Cnv_Control := "Control_DB".LCnv_Sys[4].Cnv_Level[4].Cnv1,
                 SinaSpeed := "SinaSpeed_C4104_DB",
                 ENO => #_w3);
   "C4105_FB_DB"(EN := #_w3,   // "Buffer_Conveyor_FB"
                 Cnv_Settings := "Settings_DB".LCnv_Sys[4].Cnv_Level[5].Cnv1,
                 VTD_Level := "Control_DB".VTD_Sys[4].Current_Level,
                 Safety_OK_Delayed := "Remote_Panel_DB_4".Safety_OK,
                 Safety_OK := "Remote_Panel_DB_4".Safety_Ok_Conf,
                 CNV_In_Out := "CNV_HMI".In_Out[4],
                 Cnv_Control := "Control_DB".LCnv_Sys[4].Cnv_Level[5].Cnv1,
                 SinaSpeed := "SinaSpeed_C4105_DB",
                 ENO => #_w4);
   IF #_w4 THEN
       "C4106_FB_DB"(Cnv_Settings := "Settings_DB".LCnv_Sys[4].Cnv_Level[6].Cnv1,   // "Buffer_Conveyor_FB"
                     VTD_Level := "Control_DB".VTD_Sys[4].Current_Level,
                     Safety_OK_Delayed := "Remote_Panel_DB_4".Safety_OK,
                     Safety_OK := "Remote_Panel_DB_4".Safety_Ok_Conf,
                     CNV_In_Out := "CNV_HMI".In_Out[4],
                     Cnv_Control := "Control_DB".LCnv_Sys[4].Cnv_Level[6].Cnv1,
                     SinaSpeed := "SinaSpeed_C4106_DB");
   END_IF;
   "C4107_FB_DB"(Cnv_Settings := "Settings_DB".LCnv_Sys[4].Cnv_Level[7].Cnv1,   // "Buffer_Conveyor_FB"
                 VTD_Level := "Control_DB".VTD_Sys[4].Current_Level,
                 Safety_OK_Delayed := "Remote_Panel_DB_4".Safety_OK,
                 Safety_OK := "Remote_Panel_DB_4".Safety_Ok_Conf,
                 CNV_In_Out := "CNV_HMI".In_Out[4],
                 Cnv_Control := "Control_DB".LCnv_Sys[4].Cnv_Level[7].Cnv1,
                 SinaSpeed := "SinaSpeed_C4107_DB",
                 ENO => #_w5);
   IF #_w5 THEN
       "C4108_FB_DB"(Cnv_Settings := "Settings_DB".LCnv_Sys[4].Cnv_Level[8].Cnv1,   // "Buffer_Conveyor_FB"
                     VTD_Level := "Control_DB".VTD_Sys[4].Current_Level,
                     Safety_OK_Delayed := "Remote_Panel_DB_4".Safety_OK,
                     Safety_OK := "Remote_Panel_DB_4".Safety_Ok_Conf,
                     CNV_In_Out := "CNV_HMI".In_Out[4],
                     Cnv_Control := "Control_DB".LCnv_Sys[4].Cnv_Level[8].Cnv1,
                     SinaSpeed := "SinaSpeed_C4108_DB");
   END_IF;
END_REGION

REGION Network 36: SAFETY STOPPERS Tower 1 - SYSTEM 4
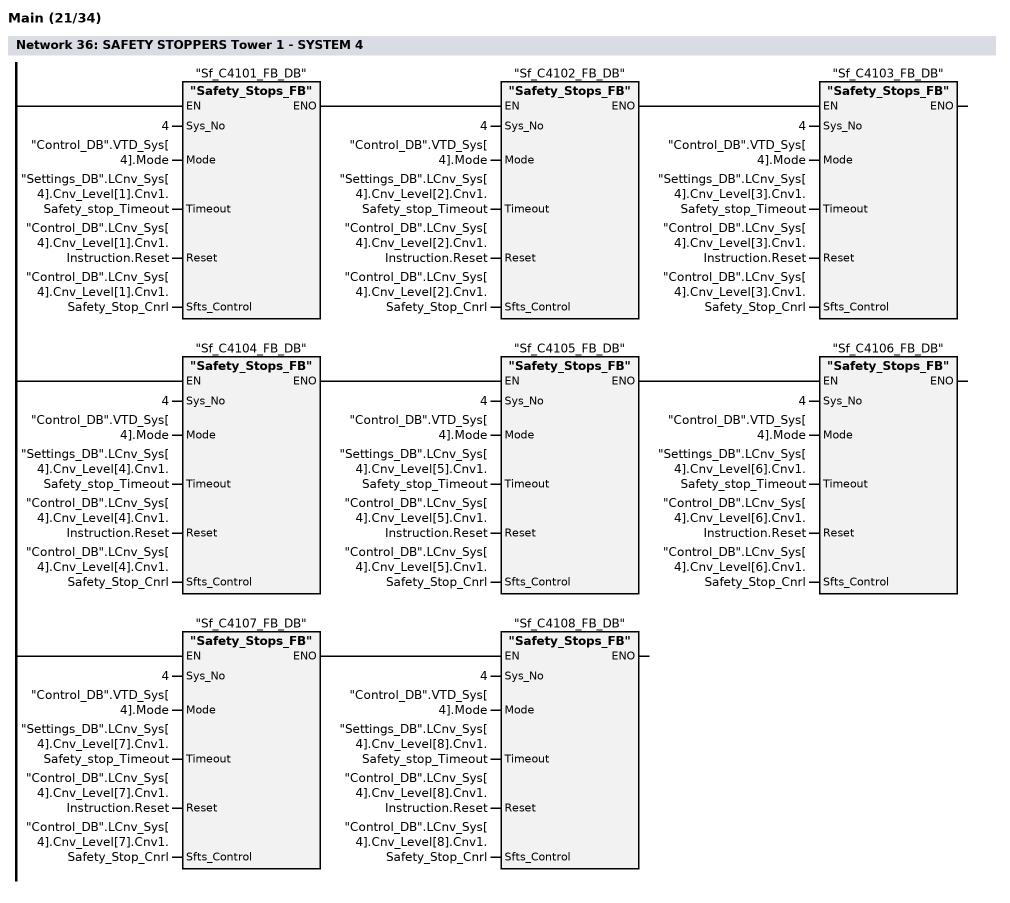
   RUNG wire#powerrail
      "Sf_C4101_FB_DB"(Sys_No := 4, Mode := "Control_DB".VTD_Sys[4].Mode, Timeout := "Settings_DB".LCnv_Sys[4].Cnv_Level[1].Cnv1.Safety_stop_Timeout, Reset := "Control_DB".LCnv_Sys[4].Cnv_Level[1].Cnv1.Instruction.Reset, Sfts_Control := "Control_DB".LCnv_Sys[4].Cnv_Level[1].Cnv1.Safety_Stop_Cnrl)
      "Sf_C4102_FB_DB"(Sys_No := 4, Mode := "Control_DB".VTD_Sys[4].Mode, Timeout := "Settings_DB".LCnv_Sys[4].Cnv_Level[2].Cnv1.Safety_stop_Timeout, Reset := "Control_DB".LCnv_Sys[4].Cnv_Level[2].Cnv1.Instruction.Reset, Sfts_Control := "Control_DB".LCnv_Sys[4].Cnv_Level[2].Cnv1.Safety_Stop_Cnrl)
      "Sf_C4103_FB_DB"(Sys_No := 4, Mode := "Control_DB".VTD_Sys[4].Mode, Timeout := "Settings_DB".LCnv_Sys[4].Cnv_Level[3].Cnv1.Safety_stop_Timeout, Reset := "Control_DB".LCnv_Sys[4].Cnv_Level[3].Cnv1.Instruction.Reset, Sfts_Control := "Control_DB".LCnv_Sys[4].Cnv_Level[3].Cnv1.Safety_Stop_Cnrl)
   END_RUNG
   RUNG wire#powerrail
      "Sf_C4104_FB_DB"(Sys_No := 4, Mode := "Control_DB".VTD_Sys[4].Mode, Timeout := "Settings_DB".LCnv_Sys[4].Cnv_Level[4].Cnv1.Safety_stop_Timeout, Reset := "Control_DB".LCnv_Sys[4].Cnv_Level[4].Cnv1.Instruction.Reset, Sfts_Control := "Control_DB".LCnv_Sys[4].Cnv_Level[4].Cnv1.Safety_Stop_Cnrl)
      "Sf_C4105_FB_DB"(Sys_No := 4, Mode := "Control_DB".VTD_Sys[4].Mode, Timeout := "Settings_DB".LCnv_Sys[4].Cnv_Level[5].Cnv1.Safety_stop_Timeout, Reset := "Control_DB".LCnv_Sys[4].Cnv_Level[5].Cnv1.Instruction.Reset, Sfts_Control := "Control_DB".LCnv_Sys[4].Cnv_Level[5].Cnv1.Safety_Stop_Cnrl)
      "Sf_C4106_FB_DB"(Sys_No := 4, Mode := "Control_DB".VTD_Sys[4].Mode, Timeout := "Settings_DB".LCnv_Sys[4].Cnv_Level[6].Cnv1.Safety_stop_Timeout, Reset := "Control_DB".LCnv_Sys[4].Cnv_Level[6].Cnv1.Instruction.Reset, Sfts_Control := "Control_DB".LCnv_Sys[4].Cnv_Level[6].Cnv1.Safety_Stop_Cnrl)
   END_RUNG
   RUNG wire#powerrail
      "Sf_C4107_FB_DB"(Sys_No := 4, Mode := "Control_DB".VTD_Sys[4].Mode, Timeout := "Settings_DB".LCnv_Sys[4].Cnv_Level[7].Cnv1.Safety_stop_Timeout, Reset := "Control_DB".LCnv_Sys[4].Cnv_Level[7].Cnv1.Instruction.Reset, Sfts_Control := "Control_DB".LCnv_Sys[4].Cnv_Level[7].Cnv1.Safety_Stop_Cnrl)
      "Sf_C4108_FB_DB"(Sys_No := 4, Mode := "Control_DB".VTD_Sys[4].Mode, Timeout := "Settings_DB".LCnv_Sys[4].Cnv_Level[8].Cnv1.Safety_stop_Timeout, Reset := "Control_DB".LCnv_Sys[4].Cnv_Level[8].Cnv1.Instruction.Reset, Sfts_Control := "Control_DB".LCnv_Sys[4].Cnv_Level[8].Cnv1.Safety_Stop_Cnrl)
   END_RUNG
   // the same network as SCL:
   "Sf_C4101_FB_DB"(Sys_No := 4,   // "Safety_Stops_FB"
                    Mode := "Control_DB".VTD_Sys[4].Mode,
                    Timeout := "Settings_DB".LCnv_Sys[4].Cnv_Level[1].Cnv1.Safety_stop_Timeout,
                    Reset := "Control_DB".LCnv_Sys[4].Cnv_Level[1].Cnv1.Instruction.Reset,
                    Sfts_Control := "Control_DB".LCnv_Sys[4].Cnv_Level[1].Cnv1.Safety_Stop_Cnrl,
                    ENO => #_w1);
   "Sf_C4102_FB_DB"(EN := #_w1,   // "Safety_Stops_FB"
                    Sys_No := 4,
                    Mode := "Control_DB".VTD_Sys[4].Mode,
                    Timeout := "Settings_DB".LCnv_Sys[4].Cnv_Level[2].Cnv1.Safety_stop_Timeout,
                    Reset := "Control_DB".LCnv_Sys[4].Cnv_Level[2].Cnv1.Instruction.Reset,
                    Sfts_Control := "Control_DB".LCnv_Sys[4].Cnv_Level[2].Cnv1.Safety_Stop_Cnrl,
                    ENO => #_w2);
   IF #_w2 THEN
       "Sf_C4103_FB_DB"(Sys_No := 4,   // "Safety_Stops_FB"
                        Mode := "Control_DB".VTD_Sys[4].Mode,
                        Timeout := "Settings_DB".LCnv_Sys[4].Cnv_Level[3].Cnv1.Safety_stop_Timeout,
                        Reset := "Control_DB".LCnv_Sys[4].Cnv_Level[3].Cnv1.Instruction.Reset,
                        Sfts_Control := "Control_DB".LCnv_Sys[4].Cnv_Level[3].Cnv1.Safety_Stop_Cnrl);
   END_IF;
   "Sf_C4104_FB_DB"(Sys_No := 4,   // "Safety_Stops_FB"
                    Mode := "Control_DB".VTD_Sys[4].Mode,
                    Timeout := "Settings_DB".LCnv_Sys[4].Cnv_Level[4].Cnv1.Safety_stop_Timeout,
                    Reset := "Control_DB".LCnv_Sys[4].Cnv_Level[4].Cnv1.Instruction.Reset,
                    Sfts_Control := "Control_DB".LCnv_Sys[4].Cnv_Level[4].Cnv1.Safety_Stop_Cnrl,
                    ENO => #_w3);
   "Sf_C4105_FB_DB"(EN := #_w3,   // "Safety_Stops_FB"
                    Sys_No := 4,
                    Mode := "Control_DB".VTD_Sys[4].Mode,
                    Timeout := "Settings_DB".LCnv_Sys[4].Cnv_Level[5].Cnv1.Safety_stop_Timeout,
                    Reset := "Control_DB".LCnv_Sys[4].Cnv_Level[5].Cnv1.Instruction.Reset,
                    Sfts_Control := "Control_DB".LCnv_Sys[4].Cnv_Level[5].Cnv1.Safety_Stop_Cnrl,
                    ENO => #_w4);
   IF #_w4 THEN
       "Sf_C4106_FB_DB"(Sys_No := 4,   // "Safety_Stops_FB"
                        Mode := "Control_DB".VTD_Sys[4].Mode,
                        Timeout := "Settings_DB".LCnv_Sys[4].Cnv_Level[6].Cnv1.Safety_stop_Timeout,
                        Reset := "Control_DB".LCnv_Sys[4].Cnv_Level[6].Cnv1.Instruction.Reset,
                        Sfts_Control := "Control_DB".LCnv_Sys[4].Cnv_Level[6].Cnv1.Safety_Stop_Cnrl);
   END_IF;
   "Sf_C4107_FB_DB"(Sys_No := 4,   // "Safety_Stops_FB"
                    Mode := "Control_DB".VTD_Sys[4].Mode,
                    Timeout := "Settings_DB".LCnv_Sys[4].Cnv_Level[7].Cnv1.Safety_stop_Timeout,
                    Reset := "Control_DB".LCnv_Sys[4].Cnv_Level[7].Cnv1.Instruction.Reset,
                    Sfts_Control := "Control_DB".LCnv_Sys[4].Cnv_Level[7].Cnv1.Safety_Stop_Cnrl,
                    ENO => #_w5);
   IF #_w5 THEN
       "Sf_C4108_FB_DB"(Sys_No := 4,   // "Safety_Stops_FB"
                        Mode := "Control_DB".VTD_Sys[4].Mode,
                        Timeout := "Settings_DB".LCnv_Sys[4].Cnv_Level[8].Cnv1.Safety_stop_Timeout,
                        Reset := "Control_DB".LCnv_Sys[4].Cnv_Level[8].Cnv1.Instruction.Reset,
                        Sfts_Control := "Control_DB".LCnv_Sys[4].Cnv_Level[8].Cnv1.Safety_Stop_Cnrl);
   END_IF;
END_REGION

REGION Network 37: SYSTEM 5
END_REGION

REGION Network 38: Level Conveyors Tower 1 - SYSTEM 5
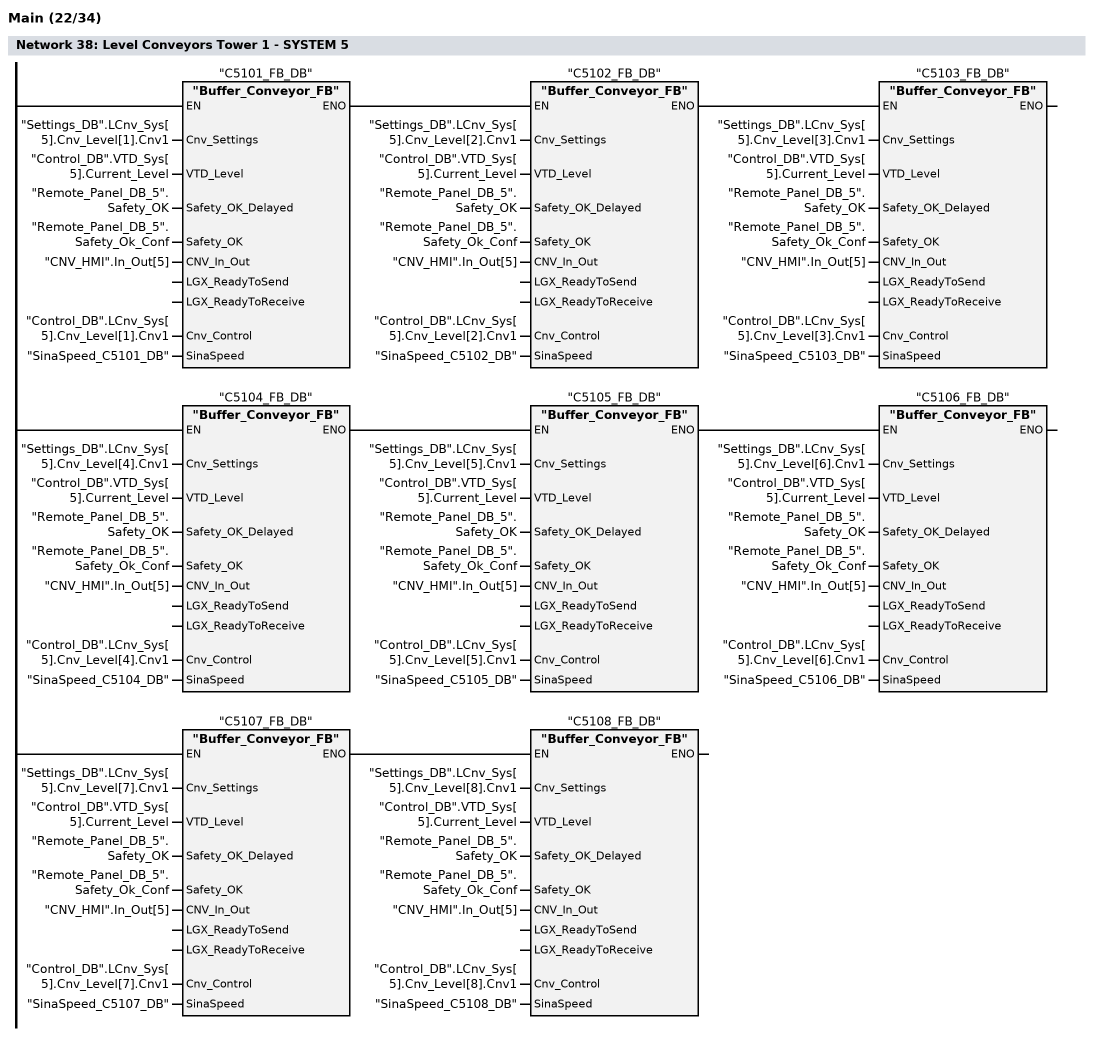
   RUNG wire#powerrail
      "C5101_FB_DB"(Cnv_Settings := "Settings_DB".LCnv_Sys[5].Cnv_Level[1].Cnv1, VTD_Level := "Control_DB".VTD_Sys[5].Current_Level, Safety_OK_Delayed := "Remote_Panel_DB_5".Safety_OK, Safety_OK := "Remote_Panel_DB_5".Safety_Ok_Conf, CNV_In_Out := "CNV_HMI".In_Out[5], LGX_ReadyToSend :=, LGX_ReadyToReceive :=, Cnv_Control := "Control_DB".LCnv_Sys[5].Cnv_Level[1].Cnv1, SinaSpeed := "SinaSpeed_C5101_DB")
      "C5102_FB_DB"(Cnv_Settings := "Settings_DB".LCnv_Sys[5].Cnv_Level[2].Cnv1, VTD_Level := "Control_DB".VTD_Sys[5].Current_Level, Safety_OK_Delayed := "Remote_Panel_DB_5".Safety_OK, Safety_OK := "Remote_Panel_DB_5".Safety_Ok_Conf, CNV_In_Out := "CNV_HMI".In_Out[5], LGX_ReadyToSend :=, LGX_ReadyToReceive :=, Cnv_Control := "Control_DB".LCnv_Sys[5].Cnv_Level[2].Cnv1, SinaSpeed := "SinaSpeed_C5102_DB")
      "C5103_FB_DB"(Cnv_Settings := "Settings_DB".LCnv_Sys[5].Cnv_Level[3].Cnv1, VTD_Level := "Control_DB".VTD_Sys[5].Current_Level, Safety_OK_Delayed := "Remote_Panel_DB_5".Safety_OK, Safety_OK := "Remote_Panel_DB_5".Safety_Ok_Conf, CNV_In_Out := "CNV_HMI".In_Out[5], LGX_ReadyToSend :=, LGX_ReadyToReceive :=, Cnv_Control := "Control_DB".LCnv_Sys[5].Cnv_Level[3].Cnv1, SinaSpeed := "SinaSpeed_C5103_DB")
   END_RUNG
   RUNG wire#powerrail
      "C5104_FB_DB"(Cnv_Settings := "Settings_DB".LCnv_Sys[5].Cnv_Level[4].Cnv1, VTD_Level := "Control_DB".VTD_Sys[5].Current_Level, Safety_OK_Delayed := "Remote_Panel_DB_5".Safety_OK, Safety_OK := "Remote_Panel_DB_5".Safety_Ok_Conf, CNV_In_Out := "CNV_HMI".In_Out[5], LGX_ReadyToSend :=, LGX_ReadyToReceive :=, Cnv_Control := "Control_DB".LCnv_Sys[5].Cnv_Level[4].Cnv1, SinaSpeed := "SinaSpeed_C5104_DB")
      "C5105_FB_DB"(Cnv_Settings := "Settings_DB".LCnv_Sys[5].Cnv_Level[5].Cnv1, VTD_Level := "Control_DB".VTD_Sys[5].Current_Level, Safety_OK_Delayed := "Remote_Panel_DB_5".Safety_OK, Safety_OK := "Remote_Panel_DB_5".Safety_Ok_Conf, CNV_In_Out := "CNV_HMI".In_Out[5], LGX_ReadyToSend :=, LGX_ReadyToReceive :=, Cnv_Control := "Control_DB".LCnv_Sys[5].Cnv_Level[5].Cnv1, SinaSpeed := "SinaSpeed_C5105_DB")
      "C5106_FB_DB"(Cnv_Settings := "Settings_DB".LCnv_Sys[5].Cnv_Level[6].Cnv1, VTD_Level := "Control_DB".VTD_Sys[5].Current_Level, Safety_OK_Delayed := "Remote_Panel_DB_5".Safety_OK, Safety_OK := "Remote_Panel_DB_5".Safety_Ok_Conf, CNV_In_Out := "CNV_HMI".In_Out[5], LGX_ReadyToSend :=, LGX_ReadyToReceive :=, Cnv_Control := "Control_DB".LCnv_Sys[5].Cnv_Level[6].Cnv1, SinaSpeed := "SinaSpeed_C5106_DB")
   END_RUNG
   RUNG wire#powerrail
      "C5107_FB_DB"(Cnv_Settings := "Settings_DB".LCnv_Sys[5].Cnv_Level[7].Cnv1, VTD_Level := "Control_DB".VTD_Sys[5].Current_Level, Safety_OK_Delayed := "Remote_Panel_DB_5".Safety_OK, Safety_OK := "Remote_Panel_DB_5".Safety_Ok_Conf, CNV_In_Out := "CNV_HMI".In_Out[5], LGX_ReadyToSend :=, LGX_ReadyToReceive :=, Cnv_Control := "Control_DB".LCnv_Sys[5].Cnv_Level[7].Cnv1, SinaSpeed := "SinaSpeed_C5107_DB")
      "C5108_FB_DB"(Cnv_Settings := "Settings_DB".LCnv_Sys[5].Cnv_Level[8].Cnv1, VTD_Level := "Control_DB".VTD_Sys[5].Current_Level, Safety_OK_Delayed := "Remote_Panel_DB_5".Safety_OK, Safety_OK := "Remote_Panel_DB_5".Safety_Ok_Conf, CNV_In_Out := "CNV_HMI".In_Out[5], LGX_ReadyToSend :=, LGX_ReadyToReceive :=, Cnv_Control := "Control_DB".LCnv_Sys[5].Cnv_Level[8].Cnv1, SinaSpeed := "SinaSpeed_C5108_DB")
   END_RUNG
   // the same network as SCL:
   "C5101_FB_DB"(Cnv_Settings := "Settings_DB".LCnv_Sys[5].Cnv_Level[1].Cnv1,   // "Buffer_Conveyor_FB"
                 VTD_Level := "Control_DB".VTD_Sys[5].Current_Level,
                 Safety_OK_Delayed := "Remote_Panel_DB_5".Safety_OK,
                 Safety_OK := "Remote_Panel_DB_5".Safety_Ok_Conf,
                 CNV_In_Out := "CNV_HMI".In_Out[5],
                 Cnv_Control := "Control_DB".LCnv_Sys[5].Cnv_Level[1].Cnv1,
                 SinaSpeed := "SinaSpeed_C5101_DB",
                 ENO => #_w1);
   "C5102_FB_DB"(EN := #_w1,   // "Buffer_Conveyor_FB"
                 Cnv_Settings := "Settings_DB".LCnv_Sys[5].Cnv_Level[2].Cnv1,
                 VTD_Level := "Control_DB".VTD_Sys[5].Current_Level,
                 Safety_OK_Delayed := "Remote_Panel_DB_5".Safety_OK,
                 Safety_OK := "Remote_Panel_DB_5".Safety_Ok_Conf,
                 CNV_In_Out := "CNV_HMI".In_Out[5],
                 Cnv_Control := "Control_DB".LCnv_Sys[5].Cnv_Level[2].Cnv1,
                 SinaSpeed := "SinaSpeed_C5102_DB",
                 ENO => #_w2);
   IF #_w2 THEN
       "C5103_FB_DB"(Cnv_Settings := "Settings_DB".LCnv_Sys[5].Cnv_Level[3].Cnv1,   // "Buffer_Conveyor_FB"
                     VTD_Level := "Control_DB".VTD_Sys[5].Current_Level,
                     Safety_OK_Delayed := "Remote_Panel_DB_5".Safety_OK,
                     Safety_OK := "Remote_Panel_DB_5".Safety_Ok_Conf,
                     CNV_In_Out := "CNV_HMI".In_Out[5],
                     Cnv_Control := "Control_DB".LCnv_Sys[5].Cnv_Level[3].Cnv1,
                     SinaSpeed := "SinaSpeed_C5103_DB");
   END_IF;
   "C5104_FB_DB"(Cnv_Settings := "Settings_DB".LCnv_Sys[5].Cnv_Level[4].Cnv1,   // "Buffer_Conveyor_FB"
                 VTD_Level := "Control_DB".VTD_Sys[5].Current_Level,
                 Safety_OK_Delayed := "Remote_Panel_DB_5".Safety_OK,
                 Safety_OK := "Remote_Panel_DB_5".Safety_Ok_Conf,
                 CNV_In_Out := "CNV_HMI".In_Out[5],
                 Cnv_Control := "Control_DB".LCnv_Sys[5].Cnv_Level[4].Cnv1,
                 SinaSpeed := "SinaSpeed_C5104_DB",
                 ENO => #_w3);
   "C5105_FB_DB"(EN := #_w3,   // "Buffer_Conveyor_FB"
                 Cnv_Settings := "Settings_DB".LCnv_Sys[5].Cnv_Level[5].Cnv1,
                 VTD_Level := "Control_DB".VTD_Sys[5].Current_Level,
                 Safety_OK_Delayed := "Remote_Panel_DB_5".Safety_OK,
                 Safety_OK := "Remote_Panel_DB_5".Safety_Ok_Conf,
                 CNV_In_Out := "CNV_HMI".In_Out[5],
                 Cnv_Control := "Control_DB".LCnv_Sys[5].Cnv_Level[5].Cnv1,
                 SinaSpeed := "SinaSpeed_C5105_DB",
                 ENO => #_w4);
   IF #_w4 THEN
       "C5106_FB_DB"(Cnv_Settings := "Settings_DB".LCnv_Sys[5].Cnv_Level[6].Cnv1,   // "Buffer_Conveyor_FB"
                     VTD_Level := "Control_DB".VTD_Sys[5].Current_Level,
                     Safety_OK_Delayed := "Remote_Panel_DB_5".Safety_OK,
                     Safety_OK := "Remote_Panel_DB_5".Safety_Ok_Conf,
                     CNV_In_Out := "CNV_HMI".In_Out[5],
                     Cnv_Control := "Control_DB".LCnv_Sys[5].Cnv_Level[6].Cnv1,
                     SinaSpeed := "SinaSpeed_C5106_DB");
   END_IF;
   "C5107_FB_DB"(Cnv_Settings := "Settings_DB".LCnv_Sys[5].Cnv_Level[7].Cnv1,   // "Buffer_Conveyor_FB"
                 VTD_Level := "Control_DB".VTD_Sys[5].Current_Level,
                 Safety_OK_Delayed := "Remote_Panel_DB_5".Safety_OK,
                 Safety_OK := "Remote_Panel_DB_5".Safety_Ok_Conf,
                 CNV_In_Out := "CNV_HMI".In_Out[5],
                 Cnv_Control := "Control_DB".LCnv_Sys[5].Cnv_Level[7].Cnv1,
                 SinaSpeed := "SinaSpeed_C5107_DB",
                 ENO => #_w5);
   IF #_w5 THEN
       "C5108_FB_DB"(Cnv_Settings := "Settings_DB".LCnv_Sys[5].Cnv_Level[8].Cnv1,   // "Buffer_Conveyor_FB"
                     VTD_Level := "Control_DB".VTD_Sys[5].Current_Level,
                     Safety_OK_Delayed := "Remote_Panel_DB_5".Safety_OK,
                     Safety_OK := "Remote_Panel_DB_5".Safety_Ok_Conf,
                     CNV_In_Out := "CNV_HMI".In_Out[5],
                     Cnv_Control := "Control_DB".LCnv_Sys[5].Cnv_Level[8].Cnv1,
                     SinaSpeed := "SinaSpeed_C5108_DB");
   END_IF;
END_REGION

REGION Network 39: SAFETY STOPPERS Tower 1 - SYSTEM 5
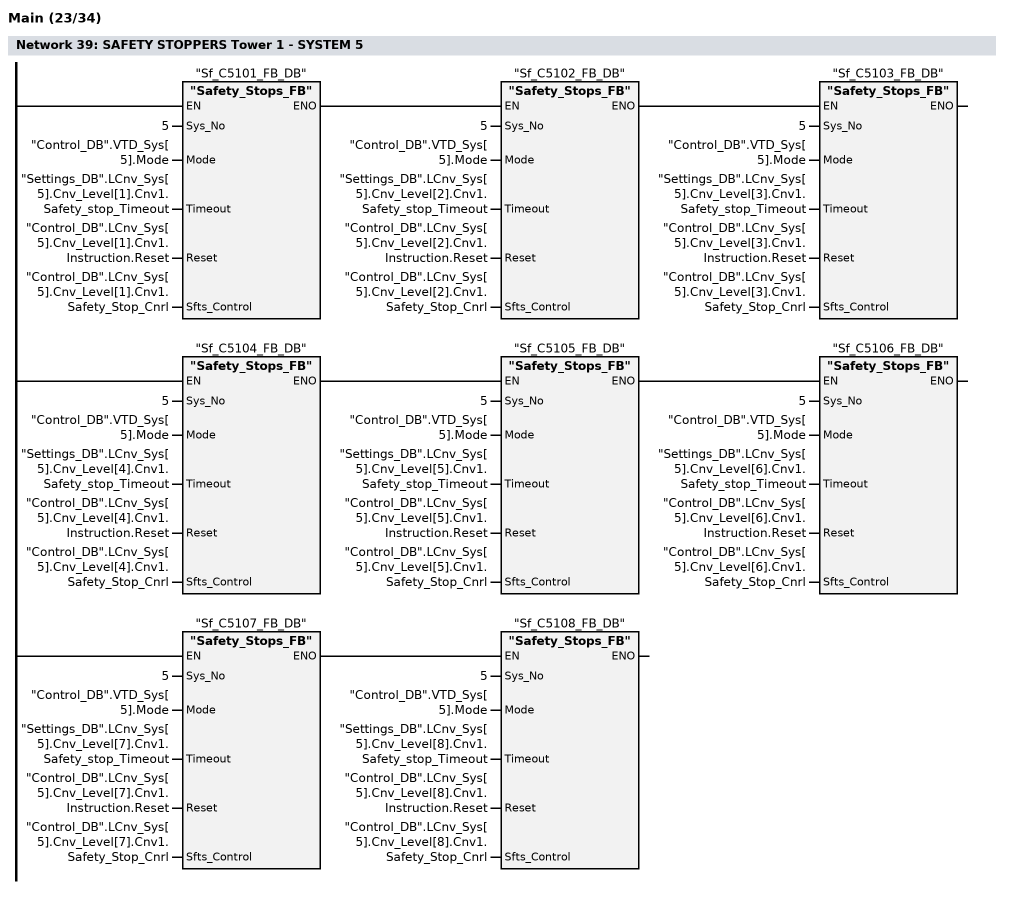
   RUNG wire#powerrail
      "Sf_C5101_FB_DB"(Sys_No := 5, Mode := "Control_DB".VTD_Sys[5].Mode, Timeout := "Settings_DB".LCnv_Sys[5].Cnv_Level[1].Cnv1.Safety_stop_Timeout, Reset := "Control_DB".LCnv_Sys[5].Cnv_Level[1].Cnv1.Instruction.Reset, Sfts_Control := "Control_DB".LCnv_Sys[5].Cnv_Level[1].Cnv1.Safety_Stop_Cnrl)
      "Sf_C5102_FB_DB"(Sys_No := 5, Mode := "Control_DB".VTD_Sys[5].Mode, Timeout := "Settings_DB".LCnv_Sys[5].Cnv_Level[2].Cnv1.Safety_stop_Timeout, Reset := "Control_DB".LCnv_Sys[5].Cnv_Level[2].Cnv1.Instruction.Reset, Sfts_Control := "Control_DB".LCnv_Sys[5].Cnv_Level[2].Cnv1.Safety_Stop_Cnrl)
      "Sf_C5103_FB_DB"(Sys_No := 5, Mode := "Control_DB".VTD_Sys[5].Mode, Timeout := "Settings_DB".LCnv_Sys[5].Cnv_Level[3].Cnv1.Safety_stop_Timeout, Reset := "Control_DB".LCnv_Sys[5].Cnv_Level[3].Cnv1.Instruction.Reset, Sfts_Control := "Control_DB".LCnv_Sys[5].Cnv_Level[3].Cnv1.Safety_Stop_Cnrl)
   END_RUNG
   RUNG wire#powerrail
      "Sf_C5104_FB_DB"(Sys_No := 5, Mode := "Control_DB".VTD_Sys[5].Mode, Timeout := "Settings_DB".LCnv_Sys[5].Cnv_Level[4].Cnv1.Safety_stop_Timeout, Reset := "Control_DB".LCnv_Sys[5].Cnv_Level[4].Cnv1.Instruction.Reset, Sfts_Control := "Control_DB".LCnv_Sys[5].Cnv_Level[4].Cnv1.Safety_Stop_Cnrl)
      "Sf_C5105_FB_DB"(Sys_No := 5, Mode := "Control_DB".VTD_Sys[5].Mode, Timeout := "Settings_DB".LCnv_Sys[5].Cnv_Level[5].Cnv1.Safety_stop_Timeout, Reset := "Control_DB".LCnv_Sys[5].Cnv_Level[5].Cnv1.Instruction.Reset, Sfts_Control := "Control_DB".LCnv_Sys[5].Cnv_Level[5].Cnv1.Safety_Stop_Cnrl)
      "Sf_C5106_FB_DB"(Sys_No := 5, Mode := "Control_DB".VTD_Sys[5].Mode, Timeout := "Settings_DB".LCnv_Sys[5].Cnv_Level[6].Cnv1.Safety_stop_Timeout, Reset := "Control_DB".LCnv_Sys[5].Cnv_Level[6].Cnv1.Instruction.Reset, Sfts_Control := "Control_DB".LCnv_Sys[5].Cnv_Level[6].Cnv1.Safety_Stop_Cnrl)
   END_RUNG
   RUNG wire#powerrail
      "Sf_C5107_FB_DB"(Sys_No := 5, Mode := "Control_DB".VTD_Sys[5].Mode, Timeout := "Settings_DB".LCnv_Sys[5].Cnv_Level[7].Cnv1.Safety_stop_Timeout, Reset := "Control_DB".LCnv_Sys[5].Cnv_Level[7].Cnv1.Instruction.Reset, Sfts_Control := "Control_DB".LCnv_Sys[5].Cnv_Level[7].Cnv1.Safety_Stop_Cnrl)
      "Sf_C5108_FB_DB"(Sys_No := 5, Mode := "Control_DB".VTD_Sys[5].Mode, Timeout := "Settings_DB".LCnv_Sys[5].Cnv_Level[8].Cnv1.Safety_stop_Timeout, Reset := "Control_DB".LCnv_Sys[5].Cnv_Level[8].Cnv1.Instruction.Reset, Sfts_Control := "Control_DB".LCnv_Sys[5].Cnv_Level[8].Cnv1.Safety_Stop_Cnrl)
   END_RUNG
   // the same network as SCL:
   "Sf_C5101_FB_DB"(Sys_No := 5,   // "Safety_Stops_FB"
                    Mode := "Control_DB".VTD_Sys[5].Mode,
                    Timeout := "Settings_DB".LCnv_Sys[5].Cnv_Level[1].Cnv1.Safety_stop_Timeout,
                    Reset := "Control_DB".LCnv_Sys[5].Cnv_Level[1].Cnv1.Instruction.Reset,
                    Sfts_Control := "Control_DB".LCnv_Sys[5].Cnv_Level[1].Cnv1.Safety_Stop_Cnrl,
                    ENO => #_w1);
   "Sf_C5102_FB_DB"(EN := #_w1,   // "Safety_Stops_FB"
                    Sys_No := 5,
                    Mode := "Control_DB".VTD_Sys[5].Mode,
                    Timeout := "Settings_DB".LCnv_Sys[5].Cnv_Level[2].Cnv1.Safety_stop_Timeout,
                    Reset := "Control_DB".LCnv_Sys[5].Cnv_Level[2].Cnv1.Instruction.Reset,
                    Sfts_Control := "Control_DB".LCnv_Sys[5].Cnv_Level[2].Cnv1.Safety_Stop_Cnrl,
                    ENO => #_w2);
   IF #_w2 THEN
       "Sf_C5103_FB_DB"(Sys_No := 5,   // "Safety_Stops_FB"
                        Mode := "Control_DB".VTD_Sys[5].Mode,
                        Timeout := "Settings_DB".LCnv_Sys[5].Cnv_Level[3].Cnv1.Safety_stop_Timeout,
                        Reset := "Control_DB".LCnv_Sys[5].Cnv_Level[3].Cnv1.Instruction.Reset,
                        Sfts_Control := "Control_DB".LCnv_Sys[5].Cnv_Level[3].Cnv1.Safety_Stop_Cnrl);
   END_IF;
   "Sf_C5104_FB_DB"(Sys_No := 5,   // "Safety_Stops_FB"
                    Mode := "Control_DB".VTD_Sys[5].Mode,
                    Timeout := "Settings_DB".LCnv_Sys[5].Cnv_Level[4].Cnv1.Safety_stop_Timeout,
                    Reset := "Control_DB".LCnv_Sys[5].Cnv_Level[4].Cnv1.Instruction.Reset,
                    Sfts_Control := "Control_DB".LCnv_Sys[5].Cnv_Level[4].Cnv1.Safety_Stop_Cnrl,
                    ENO => #_w3);
   "Sf_C5105_FB_DB"(EN := #_w3,   // "Safety_Stops_FB"
                    Sys_No := 5,
                    Mode := "Control_DB".VTD_Sys[5].Mode,
                    Timeout := "Settings_DB".LCnv_Sys[5].Cnv_Level[5].Cnv1.Safety_stop_Timeout,
                    Reset := "Control_DB".LCnv_Sys[5].Cnv_Level[5].Cnv1.Instruction.Reset,
                    Sfts_Control := "Control_DB".LCnv_Sys[5].Cnv_Level[5].Cnv1.Safety_Stop_Cnrl,
                    ENO => #_w4);
   IF #_w4 THEN
       "Sf_C5106_FB_DB"(Sys_No := 5,   // "Safety_Stops_FB"
                        Mode := "Control_DB".VTD_Sys[5].Mode,
                        Timeout := "Settings_DB".LCnv_Sys[5].Cnv_Level[6].Cnv1.Safety_stop_Timeout,
                        Reset := "Control_DB".LCnv_Sys[5].Cnv_Level[6].Cnv1.Instruction.Reset,
                        Sfts_Control := "Control_DB".LCnv_Sys[5].Cnv_Level[6].Cnv1.Safety_Stop_Cnrl);
   END_IF;
   "Sf_C5107_FB_DB"(Sys_No := 5,   // "Safety_Stops_FB"
                    Mode := "Control_DB".VTD_Sys[5].Mode,
                    Timeout := "Settings_DB".LCnv_Sys[5].Cnv_Level[7].Cnv1.Safety_stop_Timeout,
                    Reset := "Control_DB".LCnv_Sys[5].Cnv_Level[7].Cnv1.Instruction.Reset,
                    Sfts_Control := "Control_DB".LCnv_Sys[5].Cnv_Level[7].Cnv1.Safety_Stop_Cnrl,
                    ENO => #_w5);
   IF #_w5 THEN
       "Sf_C5108_FB_DB"(Sys_No := 5,   // "Safety_Stops_FB"
                        Mode := "Control_DB".VTD_Sys[5].Mode,
                        Timeout := "Settings_DB".LCnv_Sys[5].Cnv_Level[8].Cnv1.Safety_stop_Timeout,
                        Reset := "Control_DB".LCnv_Sys[5].Cnv_Level[8].Cnv1.Instruction.Reset,
                        Sfts_Control := "Control_DB".LCnv_Sys[5].Cnv_Level[8].Cnv1.Safety_Stop_Cnrl);
   END_IF;
END_REGION

REGION Network 40: Light bars
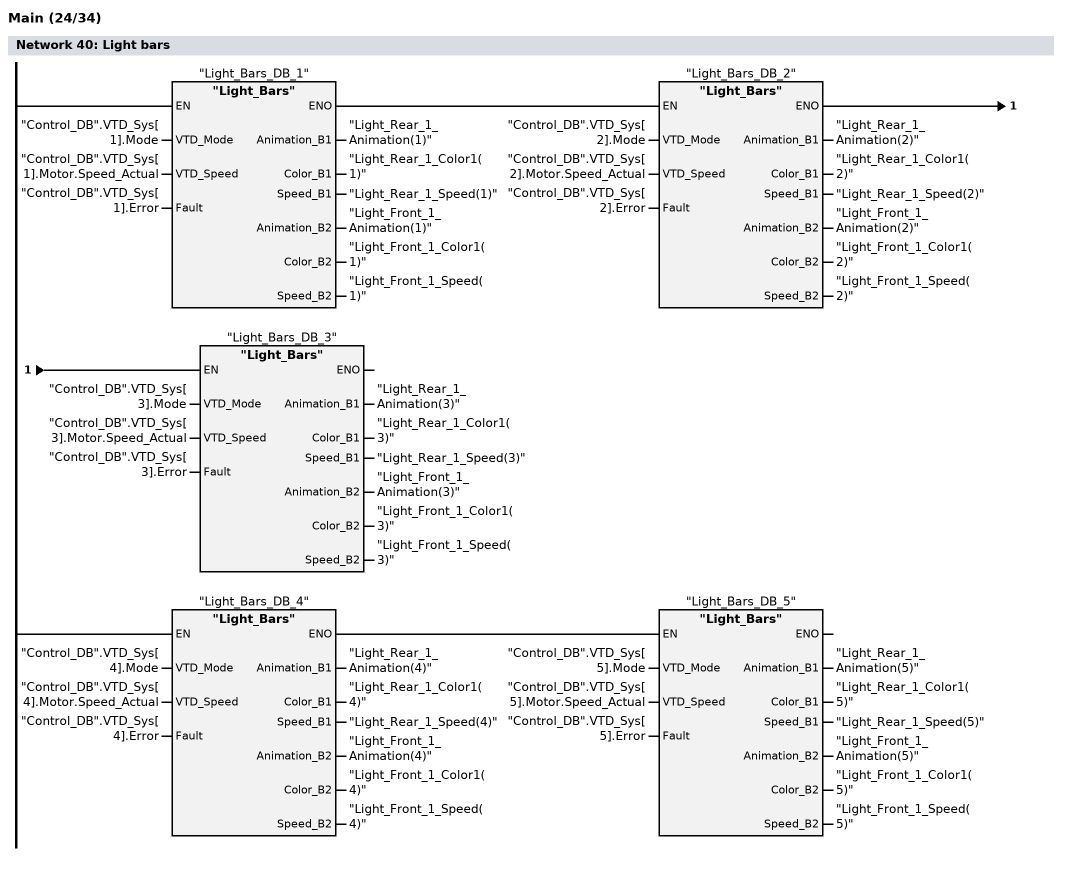
   RUNG wire#powerrail
      "Light_Bars_DB_1"(VTD_Mode := "Control_DB".VTD_Sys[1].Mode, VTD_Speed := "Control_DB".VTD_Sys[1].Motor.Speed_Actual, Fault := "Control_DB".VTD_Sys[1].Error, Animation_B1 => "Light_Rear_1_Animation(1)", Color_B1 => "Light_Rear_1_Color1(1)", Speed_B1 => "Light_Rear_1_Speed(1)", Animation_B2 => "Light_Front_1_Animation(1)", Color_B2 => "Light_Front_1_Color1(1)", Speed_B2 => "Light_Front_1_Speed(1)")
      "Light_Bars_DB_2"(VTD_Mode := "Control_DB".VTD_Sys[2].Mode, VTD_Speed := "Control_DB".VTD_Sys[2].Motor.Speed_Actual, Fault := "Control_DB".VTD_Sys[2].Error, Animation_B1 => "Light_Rear_1_Animation(2)", Color_B1 => "Light_Rear_1_Color1(2)", Speed_B1 => "Light_Rear_1_Speed(2)", Animation_B2 => "Light_Front_1_Animation(2)", Color_B2 => "Light_Front_1_Color1(2)", Speed_B2 => "Light_Front_1_Speed(2)")
      "Light_Bars_DB_3"(VTD_Mode := "Control_DB".VTD_Sys[3].Mode, VTD_Speed := "Control_DB".VTD_Sys[3].Motor.Speed_Actual, Fault := "Control_DB".VTD_Sys[3].Error, Animation_B1 => "Light_Rear_1_Animation(3)", Color_B1 => "Light_Rear_1_Color1(3)", Speed_B1 => "Light_Rear_1_Speed(3)", Animation_B2 => "Light_Front_1_Animation(3)", Color_B2 => "Light_Front_1_Color1(3)", Speed_B2 => "Light_Front_1_Speed(3)")
   END_RUNG
   RUNG wire#powerrail
      "Light_Bars_DB_4"(VTD_Mode := "Control_DB".VTD_Sys[4].Mode, VTD_Speed := "Control_DB".VTD_Sys[4].Motor.Speed_Actual, Fault := "Control_DB".VTD_Sys[4].Error, Animation_B1 => "Light_Rear_1_Animation(4)", Color_B1 => "Light_Rear_1_Color1(4)", Speed_B1 => "Light_Rear_1_Speed(4)", Animation_B2 => "Light_Front_1_Animation(4)", Color_B2 => "Light_Front_1_Color1(4)", Speed_B2 => "Light_Front_1_Speed(4)")
      "Light_Bars_DB_5"(VTD_Mode := "Control_DB".VTD_Sys[5].Mode, VTD_Speed := "Control_DB".VTD_Sys[5].Motor.Speed_Actual, Fault := "Control_DB".VTD_Sys[5].Error, Animation_B1 => "Light_Rear_1_Animation(5)", Color_B1 => "Light_Rear_1_Color1(5)", Speed_B1 => "Light_Rear_1_Speed(5)", Animation_B2 => "Light_Front_1_Animation(5)", Color_B2 => "Light_Front_1_Color1(5)", Speed_B2 => "Light_Front_1_Speed(5)")
   END_RUNG
   // the same network as SCL:
   "Light_Bars_DB_1"(VTD_Mode := "Control_DB".VTD_Sys[1].Mode,   // "Light_Bars"
                     VTD_Speed := "Control_DB".VTD_Sys[1].Motor.Speed_Actual,
                     Fault := "Control_DB".VTD_Sys[1].Error,
                     Animation_B1 => "Light_Rear_1_Animation(1)",
                     Color_B1 => "Light_Rear_1_Color1(1)",
                     Speed_B1 => "Light_Rear_1_Speed(1)",
                     Animation_B2 => "Light_Front_1_Animation(1)",
                     Color_B2 => "Light_Front_1_Color1(1)",
                     Speed_B2 => "Light_Front_1_Speed(1)",
                     ENO => #_w1);
   "Light_Bars_DB_2"(EN := #_w1,   // "Light_Bars"
                     VTD_Mode := "Control_DB".VTD_Sys[2].Mode,
                     VTD_Speed := "Control_DB".VTD_Sys[2].Motor.Speed_Actual,
                     Fault := "Control_DB".VTD_Sys[2].Error,
                     Animation_B1 => "Light_Rear_1_Animation(2)",
                     Color_B1 => "Light_Rear_1_Color1(2)",
                     Speed_B1 => "Light_Rear_1_Speed(2)",
                     Animation_B2 => "Light_Front_1_Animation(2)",
                     Color_B2 => "Light_Front_1_Color1(2)",
                     Speed_B2 => "Light_Front_1_Speed(2)",
                     ENO => #_w2);
   IF #_w2 THEN
       "Light_Bars_DB_3"(VTD_Mode := "Control_DB".VTD_Sys[3].Mode,   // "Light_Bars"
                         VTD_Speed := "Control_DB".VTD_Sys[3].Motor.Speed_Actual,
                         Fault := "Control_DB".VTD_Sys[3].Error,
                         Animation_B1 => "Light_Rear_1_Animation(3)",
                         Color_B1 => "Light_Rear_1_Color1(3)",
                         Speed_B1 => "Light_Rear_1_Speed(3)",
                         Animation_B2 => "Light_Front_1_Animation(3)",
                         Color_B2 => "Light_Front_1_Color1(3)",
                         Speed_B2 => "Light_Front_1_Speed(3)");
   END_IF;
   "Light_Bars_DB_4"(VTD_Mode := "Control_DB".VTD_Sys[4].Mode,   // "Light_Bars"
                     VTD_Speed := "Control_DB".VTD_Sys[4].Motor.Speed_Actual,
                     Fault := "Control_DB".VTD_Sys[4].Error,
                     Animation_B1 => "Light_Rear_1_Animation(4)",
                     Color_B1 => "Light_Rear_1_Color1(4)",
                     Speed_B1 => "Light_Rear_1_Speed(4)",
                     Animation_B2 => "Light_Front_1_Animation(4)",
                     Color_B2 => "Light_Front_1_Color1(4)",
                     Speed_B2 => "Light_Front_1_Speed(4)",
                     ENO => #_w3);
   IF #_w3 THEN
       "Light_Bars_DB_5"(VTD_Mode := "Control_DB".VTD_Sys[5].Mode,   // "Light_Bars"
                         VTD_Speed := "Control_DB".VTD_Sys[5].Motor.Speed_Actual,
                         Fault := "Control_DB".VTD_Sys[5].Error,
                         Animation_B1 => "Light_Rear_1_Animation(5)",
                         Color_B1 => "Light_Rear_1_Color1(5)",
                         Speed_B1 => "Light_Rear_1_Speed(5)",
                         Animation_B2 => "Light_Front_1_Animation(5)",
                         Color_B2 => "Light_Front_1_Color1(5)",
                         Speed_B2 => "Light_Front_1_Speed(5)");
   END_IF;
END_REGION

REGION Network 41: Barcode - System 1
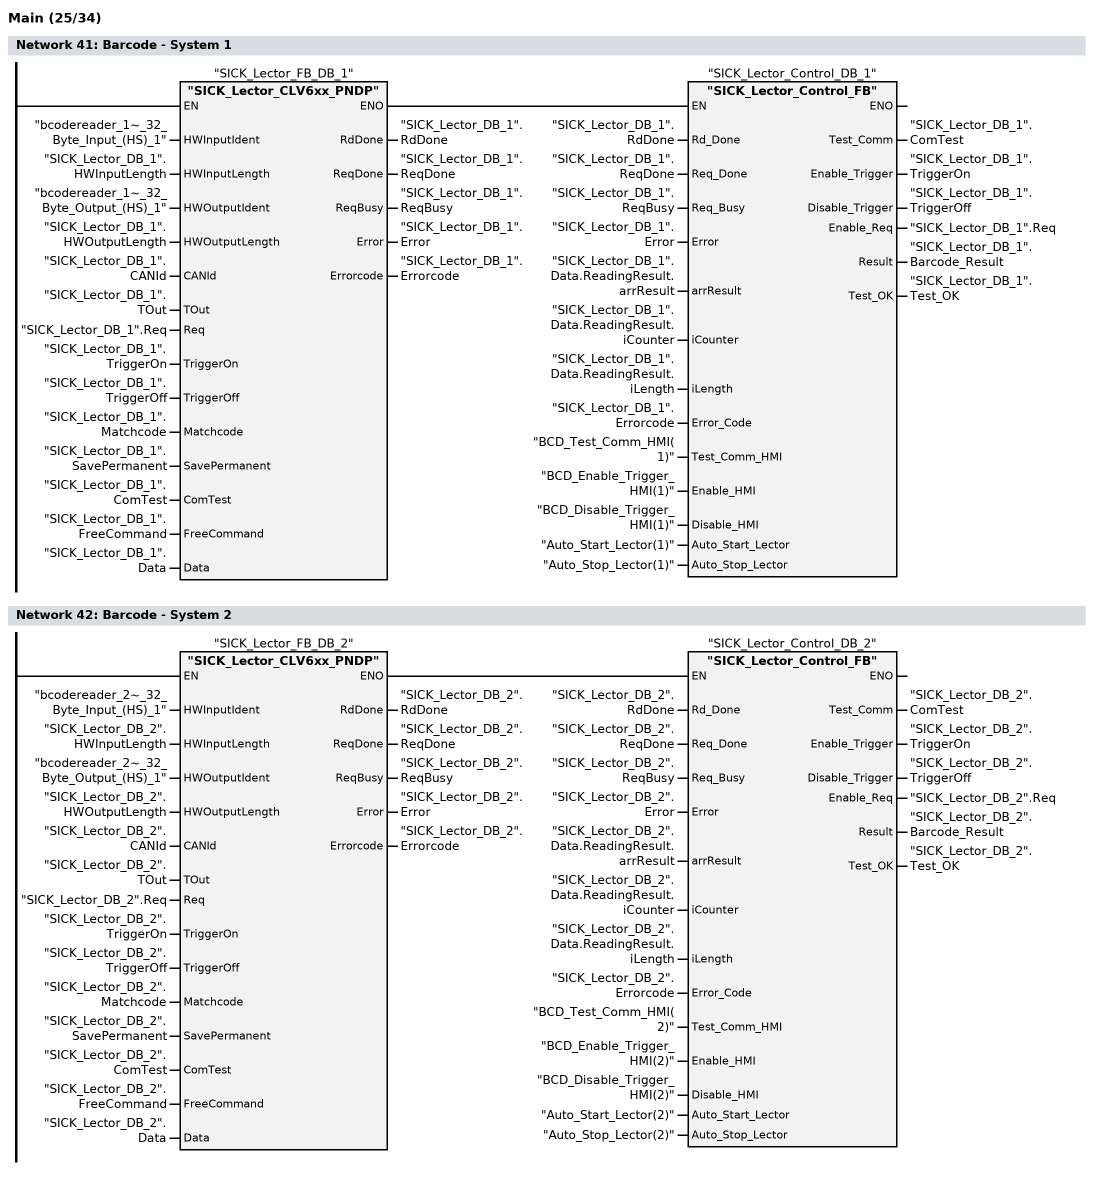
   RUNG wire#powerrail
      "SICK_Lector_FB_DB_1"(HWInputIdent := "bcodereader_1~_32_Byte_Input_(HS)_1", HWInputLength := "SICK_Lector_DB_1".HWInputLength, HWOutputIdent := "bcodereader_1~_32_Byte_Output_(HS)_1", HWOutputLength := "SICK_Lector_DB_1".HWOutputLength, CANId := "SICK_Lector_DB_1".CANId, TOut := "SICK_Lector_DB_1".TOut, Req := "SICK_Lector_DB_1".Req, TriggerOn := "SICK_Lector_DB_1".TriggerOn, TriggerOff := "SICK_Lector_DB_1".TriggerOff, Matchcode := "SICK_Lector_DB_1".Matchcode, SavePermanent := "SICK_Lector_DB_1".SavePermanent, ComTest := "SICK_Lector_DB_1".ComTest, FreeCommand := "SICK_Lector_DB_1".FreeCommand, Data := "SICK_Lector_DB_1".Data, RdDone => "SICK_Lector_DB_1".RdDone, ReqDone => "SICK_Lector_DB_1".ReqDone, ReqBusy => "SICK_Lector_DB_1".ReqBusy, Error => "SICK_Lector_DB_1".Error, Errorcode => "SICK_Lector_DB_1".Errorcode)
      "SICK_Lector_Control_DB_1"(Rd_Done := "SICK_Lector_DB_1".RdDone, Req_Done := "SICK_Lector_DB_1".ReqDone, Req_Busy := "SICK_Lector_DB_1".ReqBusy, Error := "SICK_Lector_DB_1".Error, arrResult := "SICK_Lector_DB_1".Data.ReadingResult.arrResult, iCounter := "SICK_Lector_DB_1".Data.ReadingResult.iCounter, iLength := "SICK_Lector_DB_1".Data.ReadingResult.iLength, Error_Code := "SICK_Lector_DB_1".Errorcode, Test_Comm_HMI := "BCD_Test_Comm_HMI(1)", Enable_HMI := "BCD_Enable_Trigger_HMI(1)", Disable_HMI := "BCD_Disable_Trigger_HMI(1)", Auto_Start_Lector := "Auto_Start_Lector(1)", Auto_Stop_Lector := "Auto_Stop_Lector(1)", Test_Comm => "SICK_Lector_DB_1".ComTest, Enable_Trigger => "SICK_Lector_DB_1".TriggerOn, Disable_Trigger => "SICK_Lector_DB_1".TriggerOff, Enable_Req => "SICK_Lector_DB_1".Req, Result => "SICK_Lector_DB_1".Barcode_Result, Test_OK => "SICK_Lector_DB_1".Test_OK)
   END_RUNG
   // the same network as SCL:
   "SICK_Lector_FB_DB_1"(HWInputIdent := "bcodereader_1~_32_Byte_Input_(HS)_1",   // "SICK_Lector_CLV6xx_PNDP"
                         HWInputLength := "SICK_Lector_DB_1".HWInputLength,
                         HWOutputIdent := "bcodereader_1~_32_Byte_Output_(HS)_1",
                         HWOutputLength := "SICK_Lector_DB_1".HWOutputLength,
                         CANId := "SICK_Lector_DB_1".CANId,
                         TOut := "SICK_Lector_DB_1".TOut,
                         Req := "SICK_Lector_DB_1".Req,
                         TriggerOn := "SICK_Lector_DB_1".TriggerOn,
                         TriggerOff := "SICK_Lector_DB_1".TriggerOff,
                         Matchcode := "SICK_Lector_DB_1".Matchcode,
                         SavePermanent := "SICK_Lector_DB_1".SavePermanent,
                         ComTest := "SICK_Lector_DB_1".ComTest,
                         FreeCommand := "SICK_Lector_DB_1".FreeCommand,
                         Data := "SICK_Lector_DB_1".Data,
                         RdDone => "SICK_Lector_DB_1".RdDone,
                         ReqDone => "SICK_Lector_DB_1".ReqDone,
                         ReqBusy => "SICK_Lector_DB_1".ReqBusy,
                         Error => "SICK_Lector_DB_1".Error,
                         Errorcode => "SICK_Lector_DB_1".Errorcode,
                         ENO => #_w1);
   IF #_w1 THEN
       "SICK_Lector_Control_DB_1"(Rd_Done := "SICK_Lector_DB_1".RdDone,   // "SICK_Lector_Control_FB"
                               Req_Done := "SICK_Lector_DB_1".ReqDone,
                               Req_Busy := "SICK_Lector_DB_1".ReqBusy,
                               Error := "SICK_Lector_DB_1".Error,
                               arrResult := "SICK_Lector_DB_1".Data.ReadingResult.arrResult,
                               iCounter := "SICK_Lector_DB_1".Data.ReadingResult.iCounter,
                               iLength := "SICK_Lector_DB_1".Data.ReadingResult.iLength,
                               Error_Code := "SICK_Lector_DB_1".Errorcode,
                               Test_Comm_HMI := "BCD_Test_Comm_HMI(1)",
                               Enable_HMI := "BCD_Enable_Trigger_HMI(1)",
                               Disable_HMI := "BCD_Disable_Trigger_HMI(1)",
                               Auto_Start_Lector := "Auto_Start_Lector(1)",
                               Auto_Stop_Lector := "Auto_Stop_Lector(1)",
                               Test_Comm => "SICK_Lector_DB_1".ComTest,
                               Enable_Trigger => "SICK_Lector_DB_1".TriggerOn,
                               Disable_Trigger => "SICK_Lector_DB_1".TriggerOff,
                               Enable_Req => "SICK_Lector_DB_1".Req,
                               Result => "SICK_Lector_DB_1".Barcode_Result,
                               Test_OK => "SICK_Lector_DB_1".Test_OK);
   END_IF;
END_REGION

REGION Network 42: Barcode - System 2
   RUNG wire#powerrail
      "SICK_Lector_FB_DB_2"(HWInputIdent := "bcodereader_2~_32_Byte_Input_(HS)_1", HWInputLength := "SICK_Lector_DB_2".HWInputLength, HWOutputIdent := "bcodereader_2~_32_Byte_Output_(HS)_1", HWOutputLength := "SICK_Lector_DB_2".HWOutputLength, CANId := "SICK_Lector_DB_2".CANId, TOut := "SICK_Lector_DB_2".TOut, Req := "SICK_Lector_DB_2".Req, TriggerOn := "SICK_Lector_DB_2".TriggerOn, TriggerOff := "SICK_Lector_DB_2".TriggerOff, Matchcode := "SICK_Lector_DB_2".Matchcode, SavePermanent := "SICK_Lector_DB_2".SavePermanent, ComTest := "SICK_Lector_DB_2".ComTest, FreeCommand := "SICK_Lector_DB_2".FreeCommand, Data := "SICK_Lector_DB_2".Data, RdDone => "SICK_Lector_DB_2".RdDone, ReqDone => "SICK_Lector_DB_2".ReqDone, ReqBusy => "SICK_Lector_DB_2".ReqBusy, Error => "SICK_Lector_DB_2".Error, Errorcode => "SICK_Lector_DB_2".Errorcode)
      "SICK_Lector_Control_DB_2"(Rd_Done := "SICK_Lector_DB_2".RdDone, Req_Done := "SICK_Lector_DB_2".ReqDone, Req_Busy := "SICK_Lector_DB_2".ReqBusy, Error := "SICK_Lector_DB_2".Error, arrResult := "SICK_Lector_DB_2".Data.ReadingResult.arrResult, iCounter := "SICK_Lector_DB_2".Data.ReadingResult.iCounter, iLength := "SICK_Lector_DB_2".Data.ReadingResult.iLength, Error_Code := "SICK_Lector_DB_2".Errorcode, Test_Comm_HMI := "BCD_Test_Comm_HMI(2)", Enable_HMI := "BCD_Enable_Trigger_HMI(2)", Disable_HMI := "BCD_Disable_Trigger_HMI(2)", Auto_Start_Lector := "Auto_Start_Lector(2)", Auto_Stop_Lector := "Auto_Stop_Lector(2)", Test_Comm => "SICK_Lector_DB_2".ComTest, Enable_Trigger => "SICK_Lector_DB_2".TriggerOn, Disable_Trigger => "SICK_Lector_DB_2".TriggerOff, Enable_Req => "SICK_Lector_DB_2".Req, Result => "SICK_Lector_DB_2".Barcode_Result, Test_OK => "SICK_Lector_DB_2".Test_OK)
   END_RUNG
   // the same network as SCL:
   "SICK_Lector_FB_DB_2"(HWInputIdent := "bcodereader_2~_32_Byte_Input_(HS)_1",   // "SICK_Lector_CLV6xx_PNDP"
                         HWInputLength := "SICK_Lector_DB_2".HWInputLength,
                         HWOutputIdent := "bcodereader_2~_32_Byte_Output_(HS)_1",
                         HWOutputLength := "SICK_Lector_DB_2".HWOutputLength,
                         CANId := "SICK_Lector_DB_2".CANId,
                         TOut := "SICK_Lector_DB_2".TOut,
                         Req := "SICK_Lector_DB_2".Req,
                         TriggerOn := "SICK_Lector_DB_2".TriggerOn,
                         TriggerOff := "SICK_Lector_DB_2".TriggerOff,
                         Matchcode := "SICK_Lector_DB_2".Matchcode,
                         SavePermanent := "SICK_Lector_DB_2".SavePermanent,
                         ComTest := "SICK_Lector_DB_2".ComTest,
                         FreeCommand := "SICK_Lector_DB_2".FreeCommand,
                         Data := "SICK_Lector_DB_2".Data,
                         RdDone => "SICK_Lector_DB_2".RdDone,
                         ReqDone => "SICK_Lector_DB_2".ReqDone,
                         ReqBusy => "SICK_Lector_DB_2".ReqBusy,
                         Error => "SICK_Lector_DB_2".Error,
                         Errorcode => "SICK_Lector_DB_2".Errorcode,
                         ENO => #_w1);
   IF #_w1 THEN
       "SICK_Lector_Control_DB_2"(Rd_Done := "SICK_Lector_DB_2".RdDone,   // "SICK_Lector_Control_FB"
                               Req_Done := "SICK_Lector_DB_2".ReqDone,
                               Req_Busy := "SICK_Lector_DB_2".ReqBusy,
                               Error := "SICK_Lector_DB_2".Error,
                               arrResult := "SICK_Lector_DB_2".Data.ReadingResult.arrResult,
                               iCounter := "SICK_Lector_DB_2".Data.ReadingResult.iCounter,
                               iLength := "SICK_Lector_DB_2".Data.ReadingResult.iLength,
                               Error_Code := "SICK_Lector_DB_2".Errorcode,
                               Test_Comm_HMI := "BCD_Test_Comm_HMI(2)",
                               Enable_HMI := "BCD_Enable_Trigger_HMI(2)",
                               Disable_HMI := "BCD_Disable_Trigger_HMI(2)",
                               Auto_Start_Lector := "Auto_Start_Lector(2)",
                               Auto_Stop_Lector := "Auto_Stop_Lector(2)",
                               Test_Comm => "SICK_Lector_DB_2".ComTest,
                               Enable_Trigger => "SICK_Lector_DB_2".TriggerOn,
                               Disable_Trigger => "SICK_Lector_DB_2".TriggerOff,
                               Enable_Req => "SICK_Lector_DB_2".Req,
                               Result => "SICK_Lector_DB_2".Barcode_Result,
                               Test_OK => "SICK_Lector_DB_2".Test_OK);
   END_IF;
END_REGION

